# B&R Automation Studio project AS_Project
Automation Studio 6.7.1.5; technology packages: OpcUaCs 6.7.0

## Configuration Config1

CPU 5APC3100.KBU2-000, AutomationRuntime 6.8.1, Build 11.3.0

### Task classes (Cpu.sw)
```
Cyclic#4:
  AltDBExamp <- AltDBExample.prg
Libraries: AltDB, AsTCP, runtime, AsBrStr
```

### Hardware
```
5APC3100_KBU2_000 : 5APC3100.KBU2-000 v2.3.1.0
  Connector IF3:
    AssignedOperatingSystem = ARemb
    ActivateDevice = 1
  Connector IF4:
    AssignedOperatingSystem = ARemb
    ActivateDevice = 1
  Connector IF5:
    AssignedOperatingSystem = ARemb
  Connector IF6:
    AssignedOperatingSystem = ARemb
  Connector IF7:
    AssignedOperatingSystem = ARemb
  Connector IF8:
    AssignedOperatingSystem = ARemb
  ConfigurationID = AltDB_Config1
  Simulation = 1
  ActivateEncryption = 0
  FileDevice1
  FileDeviceName1 = USER
  FileDevicePath1 = USER_PATH
```

### BRRole.brrole - 5APC3100_KBU2_000/AccessAndSecurity/UserRoleSystem/BRRole.brrole
```
Element BR_Anonymous (Type=BRRole)
Element BR_Engineer (Type=BRRole)
Element BR_Observer (Type=BRRole)
Element BR_SafetyAdmin (Type=BRRole)
Element BR_SecurityAdmin (Type=BRRole)
```

- Physical/Config1/5APC3100_KBU2_000/IoMap.iom: same as Physical/Config1/5APC3100_KBU2_000/Cpu.per
- Physical/Config1/5APC3100_KBU2_000/PvMap.vvm: same as Physical/Config1/5APC3100_KBU2_000/Cpu.per
- Safety project (password-protected, skipped)

## Logical view

Binary libraries used (declarations not repeated): operator, runtime, AsIecCon, AsTCP, AsBrStr

### Global.typ - Global data types
```iecst
TYPE
	ReceipeType : 	STRUCT
		price : REAL;				(*recipe price*)
		setTemp : REAL;				(*set temperature*)
		milk : REAL;				(*milk quantity*)
		sugar : REAL;				(*sugar quantity*)
		coffee : REAL;				(*coffee quantity*)
		water : REAL;				(*water quantity*)
	END_STRUCT;
	ParType : 	STRUCT
		receipe : ReceipeType;		(*active recipe parameters*)
	END_STRUCT;
	MainLogicType : 	STRUCT
		par : ParType;				(*parameter structure*)
	END_STRUCT;
END_TYPE
```

### Global.var - Global variables
```iecst
VAR
gMainLogic : MainLogicType;
END_VAR

VAR CONSTANT

END_VAR
```

### Package Logical/Libraries - Global libraries

### Library Logical/Libraries/AltDB (ANSIC, version 1.0.2)
Depends on: AsTCP

#### Types.typ - Exported data types
```iecst
TYPE
	(*Extension type (not part of AsDb): internal diagnostic snapshot of
	a connection, returned by the extension FB dbGetConnState. Exposes
	the state machine of Section 9.2 plus buffering/parsing counters so
	a stuck connection (e.g. permanently ERR_FUB_BUSY) can be diagnosed
	without reading this library's C sources.*)
	AltDBConnStateType : STRUCT
		state				: UINT;		(*CONNSTATE_*, see Priv.var - OPENING/CONNECTING/PRELOGIN/LOGIN/IDLE/EXECUTING/IN_RESULT/BROKEN/FAILED*)
		netStep				: UINT;		(*sub-state of the current network operation (0=send,1=recv)*)
		jobKind				: UINT;		(*JOB_* - which FB currently owns this connection's job, JOB_NONE if idle*)
		locked				: BOOL;		(*TRUE while a job is in progress on this connection*)
		tcpIdent			: UDINT;	(*AsTCP socket identifier, 0 = not opened yet*)
		encoding			: UINT;		(*DBENC_ISO_8859_1 (0) / DBENC_UTF_8 (1)*)
		packetSize			: UINT;		(*negotiated TDS packet size*)
		sendLen				: UDINT;	(*total bytes of the outgoing message currently being sent*)
		sendPos				: UDINT;	(*bytes already handed to TcpSend*)
		tokLen				: UDINT;	(*bytes currently buffered in the de-framed token stream*)
		tokPos				: UDINT;	(*parser read cursor into the token stream*)
		statementActive		: BOOL;		(*TRUE once dbExecuteSql has completed at least once*)
		columnCount			: INT;		(*column count of the current result set, 0 if none*)
		hasResultSet		: BOOL;		(*current statement produced a result set*)
		resultSetOpen		: BOOL;		(*result set still has rows pending / not yet exhausted*)
		rowReady			: BOOL;		(*a row is currently buffered and ready for dbGetData*)
		noMoreRows			: BOOL;		(*end of the current result set has been reached*)
		affectedRows		: UDINT;
		affectedRowsKnown	: BOOL;
		diagCount			: UINT;		(*number of diagnostic records currently in the ring*)
		diagReadIdx			: UINT;		(*index of the next unread diagnostic record*)
		serverVersion		: STRING[31];	(*"mm.mm.bbbb" once LOGINACK has been received, else empty*)
	END_STRUCT;
END_TYPE
```

#### Constants.var - Exported constants
```iecst
VAR CONSTANT
	DB_SYSTEM_SYBASE				: UINT := 1;		(*Sybase database*)
	DB_SYSTEM_MS_SQL				: UINT := 2;		(*Microsoft SQL database*)

	DB_DEFAULT_PORT					: UINT := 5000;		(*default database port*)

	DB_SQL_ERROR					: INT := -1;		(*SQL error*)
	DB_SQL_INVALID_HANDLE			: INT := -2;		(*invalid SQL database handle*)
	DB_SQL_NO_DATA					: INT := 100;		(*no data available*)

	DB_SQL_CHAR						: INT := 1;			(*character data type of either fixed length or variable length*)
	DB_SQL_NUMERIC					: INT := 2;			(*numeric data type with fixed precision and scale*)
	DB_SQL_DECIMAL					: INT := 3;			(*numeric data type with fixed precision and scale*)
	DB_SQL_BIGINT					: INT := -25;		(*big integer 8 bytes*)
	DB_SQL_INTEGER					: INT := 4;			(*DINT*)
	DB_SQL_SMALLINT					: INT := 5;			(*INT*)
	DB_SQL_TINYINT					: INT := -6;		(*SINT*)
	DB_SQL_REAL						: INT := 7;			(*REAL*)
	DB_SQL_DOUBLE					: INT := 8;			(*LREAL*)
	DB_SQL_DATE						: INT := 9;			(*date, 6 bytes: yy.mm.dd*)
	DB_SQL_TIME						: INT := 10;		(*time of a day without time zone based on a 24-hour clock, 6 bytes: hh:mm:ss*)
	DB_SQL_TIMESTAMP				: INT := 11;		(*DB_SQL_DATE + TIME 12 bytes: yy.mm.dd hh:mm:ss*)
	DB_SQL_GUID						: INT := -11;		(*16 byte GUID*)

	DB_IT_SQL_ACCESSIBLE_TABLES				: UINT := 19;		(*SQL_ACCESSIBLE_TABLES*)
	DB_IT_SQL_ACTIVE_ENVIRONMENTS			: UINT := 116;		(*SQL_ACTIVE_ENVIRONMENTS*)
	DB_IT_SQL_AGGREGATE_FUNCTIONS			: UINT := 169;		(*SQL_AGGREGATE_FUNCTIONS*)
	DB_IT_SQL_ALTER_DOMAIN					: UINT := 117;		(*SQL_ALTER_DOMAIN*)
	DB_IT_SQL_ALTER_TABLE					: UINT := 86;		(*SQL_ALTER_TABLE*)
	DB_IT_SQL_ASYNC_MODE					: UINT := 10021;		(*SQL_ASYNC_MODE*)
	DB_IT_SQL_BATCH_ROW_COUNT				: UINT := 120;		(*SQL_BATCH_ROW_COUNT*)
	DB_IT_SQL_BATCH_SUPPORT					: UINT := 121;		(*SQL_BATCH_SUPPORT*)
	DB_IT_SQL_BOOKMARK_PERSISTENCE			: UINT := 82;		(*SQL_BOOKMARK_PERSISTENCE*)
	DB_IT_SQL_CATALOG_LOCATION				: UINT := 114;		(*SQL_CATALOG_LOCATION*)
	DB_IT_SQL_CATALOG_NAME					: UINT := 10003;		(*SQL_CATALOG_NAME*)
	DB_IT_SQL_CATALOG_NAME_SEPARATOR		: UINT := 41;		(*SQL_CATALOG_NAME_SEPARATOR*)
	DB_IT_SQL_CATALOG_TERM					: UINT := 42;		(*SQL_CATALOG_TERM*)
	DB_IT_SQL_CATALOG_USAGE					: UINT := 92;		(*SQL_CATALOG_USAGE*)
	DB_IT_SQL_COLUMN_ALIAS					: UINT := 87;		(*SQL_COLUMN_ALIAS*)
	DB_IT_SQL_CONCAT_NULL_BEHAVIOR			: UINT := 22;		(*SQL_CONCAT_NULL_BEHAVIOR*)
	DB_IT_SQL_CONVERT_BINARY				: UINT := 54;		(*SQL_CONVERT_BINARY*)
	DB_IT_SQL_CONVERT_BIT					: UINT := 55;		(*SQL_CONVERT_BIT*)
	DB_IT_SQL_CONVERT_CHAR					: UINT := 56;		(*SQL_CONVERT_CHAR*)
	DB_IT_SQL_CONVERT_DECIMAL				: UINT := 58;		(*SQL_CONVERT_DECIMAL*)
	DB_IT_SQL_CONVERT_FLOAT					: UINT := 60;		(*SQL_CONVERT_FLOAT*)
	DB_IT_SQL_CONVERT_FUNCTIONS				: UINT := 48;		(*SQL_CONVERT_FUNCTIONS*)
	DB_IT_SQL_CONVERT_INTEGER				: UINT := 61;		(*SQL_CONVERT_INTEGER*)
	DB_IT_SQL_CONVERT_LONGVARBINARY			: UINT := 71;		(*SQL_CONVERT_LONGVARBINARY*)
	DB_IT_SQL_CONVERT_LONGVARCHAR			: UINT := 62;		(*SQL_CONVERT_LONGVARCHAR*)
	DB_IT_SQL_CONVERT_NUMERIC				: UINT := 63;		(*SQL_CONVERT_NUMERIC*)
	DB_IT_SQL_CONVERT_REAL					: UINT := 64;		(*SQL_CONVERT_REAL*)
	DB_IT_SQL_CONVERT_SMALLINT				: UINT := 65;		(*SQL_CONVERT_SMALLINT*)
	DB_IT_SQL_CONVERT_TIMESTAMP				: UINT := 67;		(*SQL_CONVERT_TIMESTAMP*)
	DB_IT_SQL_CONVERT_TINYINT				: UINT := 68;		(*SQL_CONVERT_TINYINT*)
	DB_IT_SQL_CONVERT_VARBINARY				: UINT := 69;		(*SQL_CONVERT_VARBINARY*)
	DB_IT_SQL_CONVERT_VARCHAR				: UINT := 70;		(*SQL_CONVERT_VARCHAR*)
	DB_IT_SQL_CONVERT_WCHAR					: UINT := 122;		(*SQL_CONVERT_WCHAR*)
	DB_IT_SQL_CONVERT_WLONGVARCHAR			: UINT := 125;		(*SQL_CONVERT_WLONGVARCHAR*)
	DB_IT_SQL_CONVERT_WVARCHAR				: UINT := 126;		(*SQL_CONVERT_WVARCHAR*)
	DB_IT_SQL_CORRELATION_NAME				: UINT := 74;		(*SQL_CORRELATION_NAME*)
	DB_IT_SQL_CREATE_ASSERTION				: UINT := 127;		(*SQL_CREATE_ASSERTION*)
	DB_IT_SQL_CREATE_CHARACTER_SET			: UINT := 128;		(*SQL_CREATE_CHARACTER_SET*)
	DB_IT_SQL_CREATE_COLLATION				: UINT := 129;		(*SQL_CREATE_COLLATION*)
	DB_IT_SQL_CREATE_DOMAIN					: UINT := 130;		(*SQL_CREATE_DOMAIN*)
	DB_IT_SQL_CREATE_SCHEMA					: UINT := 131;		(*SQL_CREATE_SCHEMA*)
	DB_IT_SQL_CREATE_TABLE					: UINT := 132;		(*SQL_CREATE_TABLE*)
	DB_IT_SQL_CREATE_TRANSLATION			: UINT := 133;		(*SQL_CREATE_TRANSLATION*)
	DB_IT_SQL_CREATE_VIEW					: UINT := 134;		(*SQL_CREATE_VIEW*)
	DB_IT_SQL_CURSOR_COMMIT_BEHAVIOR		: UINT := 23;		(*SQL_CURSOR_COMMIT_BEHAVIOR*)
	DB_IT_SQL_CURSOR_ROLLBACK_BEHAV			: UINT := 24;		(*SQL_CURSOR_ROLLBACK_BEHAVIOR*)
	DB_IT_SQL_CURSOR_SENSITIVITY			: UINT := 10001;		(*SQL_CURSOR_SENSITIVITY*)
	DB_IT_SQL_DATA_SOURCE_NAME				: UINT := 2;		(*SQL_DATA_SOURCE_NAME*)
	DB_IT_SQL_DATA_SOURCE_READ_ONLY			: UINT := 25;		(*SQL_DATA_SOURCE_READ_ONLY*)
	DB_IT_SQL_DATABASE_NAME					: UINT := 16;		(*SQL_DATABASE_NAME*)
	DB_IT_SQL_DATETIME_LITERALS				: UINT := 119;		(*SQL_DATETIME_LITERALS*)
	DB_IT_SQL_DBMS_NAME						: UINT := 17;		(*SQL_DBMS_NAME*)
	DB_IT_SQL_DBMS_VER						: UINT := 18;		(*SQL_DBMS_VER*)
	DB_IT_SQL_DDL_INDEX						: UINT := 170;		(*SQL_DDL_INDEX*)
	DB_IT_SQL_DEFAULT_TXN_ISOLATION			: UINT := 26;		(*SQL_DEFAULT_TXN_ISOLATION*)
	DB_IT_SQL_DESCRIBE_PARAMETER			: UINT := 10002;		(*SQL_DESCRIBE_PARAMETER*)
	DB_IT_SQL_DRIVER_HDBC					: UINT := 3;		(*SQL_DRIVER_HDBC*)
	DB_IT_SQL_DRIVER_HENV					: UINT := 4;		(*SQL_DRIVER_HENV*)
	DB_IT_SQL_DRIVER_HSTMT					: UINT := 5;		(*SQL_DRIVER_HSTMT*)
	DB_IT_SQL_DRIVER_NAME					: UINT := 6;		(*SQL_DRIVER_NAME*)
	DB_IT_SQL_DRIVER_ODBC_VER				: UINT := 77;		(*SQL_DRIVER_ODBC_VER*)
	DB_IT_SQL_DRIVER_VER					: UINT := 7;		(*SQL_DRIVER_VER*)
	DB_IT_SQL_DROP_ASSERTION				: UINT := 136;		(*SQL_DROP_ASSERTION*)
	DB_IT_SQL_DROP_CHARACTER_SET			: UINT := 137;		(*SQL_DROP_CHARACTER_SET*)
	DB_IT_SQL_DROP_COLLATION				: UINT := 138;		(*SQL_DROP_COLLATION*)
	DB_IT_SQL_DROP_DOMAIN					: UINT := 139;		(*SQL_DROP_DOMAIN*)
	DB_IT_SQL_DROP_SCHEMA					: UINT := 140;		(*SQL_DROP_SCHEMA*)
	DB_IT_SQL_DROP_TABLE					: UINT := 141;		(*SQL_DROP_TABLE*)
	DB_IT_SQL_DROP_TRANSLATION				: UINT := 142;		(*SQL_DROP_TRANSLATION*)
	DB_IT_SQL_DROP_VIEW						: UINT := 143;		(*SQL_DROP_VIEW*)
	DB_IT_SQL_DYNAMIC_CURSOR_ATTR1			: UINT := 144;		(*SQL_DYNAMIC_CURSOR_ATTRIBUTES1*)
	DB_IT_SQL_DYNAMIC_CURSOR_ATTR2			: UINT := 145;		(*SQL_DYNAMIC_CURSOR_ATTRIBUTES2*)
	DB_IT_SQL_EXPRESSIONS_IN_ORDERBY		: UINT := 27;		(*SQL_EXPRESSIONS_IN_ORDERBY*)
	DB_IT_SQL_FETCH_DIRECTION				: UINT := 8;		(*SQL_FETCH_DIRECTION*)
	DB_IT_SQL_FILE_USAGE					: UINT := 84;		(*SQL_FILE_USAGE*)
	DB_IT_SQL_FORW_ONLY_CURSOR_ATTR1		: UINT := 146;		(*SQL_FORWARD_ONLY_CURSOR_ATTRIBUTES1*)
	DB_IT_SQL_FORW_ONLY_CURSOR_ATTR2		: UINT := 147;		(*SQL_FORWARD_ONLY_CURSOR_ATTRIBUTES2*)
	DB_IT_SQL_GETDATA_EXTENSIONS			: UINT := 81;		(*SQL_GETDATA_EXTENSIONS*)
	DB_IT_SQL_GROUP_BY						: UINT := 88;		(*SQL_GROUP_BY*)
	DB_IT_SQL_IDENTIFIER_CASE				: UINT := 28;		(*SQL_IDENTIFIER_CASE*)
	DB_IT_SQL_IDENTIFIER_QUOTE_CHAR			: UINT := 29;		(*SQL_IDENTIFIER_QUOTE_CHAR*)
	DB_IT_SQL_INDEX_KEYWORDS				: UINT := 148;		(*SQL_INDEX_KEYWORDS*)
	DB_IT_SQL_INFO_SCHEMA_VIEWS				: UINT := 149;		(*SQL_INFO_SCHEMA_VIEWS*)
	DB_IT_SQL_INSERT_STATEMENT				: UINT := 172;		(*SQL_INSERT_STATEMENT*)
	DB_IT_SQL_INTEGRITY						: UINT := 73;		(*SQL_INTEGRITY*)
	DB_IT_SQL_KEYSET_CURSOR_ATTR1			: UINT := 150;		(*SQL_KEYSET_CURSOR_ATTRIBUTES1*)
	DB_IT_SQL_KEYSET_CURSOR_ATTR2			: UINT := 151;		(*SQL_KEYSET_CURSOR_ATTRIBUTES2*)
	DB_IT_SQL_KEYWORDS						: UINT := 89;		(*SQL_KEYWORDS*)
	DB_IT_SQL_LIKE_ESCAPE_CLAUSE			: UINT := 113;		(*SQL_LIKE_ESCAPE_CLAUSE*)
	DB_IT_SQL_LOCK_TYPES					: UINT := 78;		(*SQL_LOCK_TYPES*)
	DB_IT_SQL_MAX_ASYNC_CONCUR_STMT			: UINT := 10022;		(*SQL_MAX_ASYNC_CONCURRENT_STATEMENTS*)
	DB_IT_SQL_MAX_BINARY_LITERAL_LEN		: UINT := 112;		(*SQL_MAX_BINARY_LITERAL_LEN*)
	DB_IT_SQL_MAX_CATALOG_NAME_LEN			: UINT := 34;		(*SQL_MAX_CATALOG_NAME_LEN*)
	DB_IT_SQL_MAX_CHAR_LITERAL_LEN			: UINT := 108;		(*SQL_MAX_CHAR_LITERAL_LEN*)
	DB_IT_SQL_MAX_COLUMN_NAME_LEN			: UINT := 30;		(*SQL_MAX_COLUMN_NAME_LEN*)
	DB_IT_SQL_MAX_COLS_IN_GROUP_BY			: UINT := 97;		(*SQL_MAX_COLUMNS_IN_GROUP_BY*)
	DB_IT_SQL_MAX_COLUMNS_IN_INDEX			: UINT := 98;		(*SQL_MAX_COLUMNS_IN_INDEX*)
	DB_IT_SQL_MAX_COLS_IN_ORDER_BY			: UINT := 99;		(*SQL_MAX_COLUMNS_IN_ORDER_BY*)
	DB_IT_SQL_MAX_COLUMNS_IN_SELECT			: UINT := 100;		(*SQL_MAX_COLUMNS_IN_SELECT*)
	DB_IT_SQL_MAX_COLUMNS_IN_TABLE			: UINT := 101;		(*SQL_MAX_COLUMNS_IN_TABLE*)
	DB_IT_SQL_MAX_CONCUR_ACTIVITIES			: UINT := 1;		(*SQL_MAX_CONCURRENT_ACTIVITIES*)
	DB_IT_SQL_MAX_CURSOR_NAME_LEN			: UINT := 31;		(*SQL_MAX_CURSOR_NAME_LEN*)
	DB_IT_SQL_MAX_DRIVER_CONNECTIONS		: UINT := 0;		(*SQL_MAX_DRIVER_CONNECTIONS*)
	DB_IT_SQL_MAX_IDENTIFIER_LEN			: UINT := 10005;		(*SQL_MAX_IDENTIFIER_LEN*)
	DB_IT_SQL_MAX_INDEX_SIZE				: UINT := 102;		(*SQL_MAX_INDEX_SIZE*)
	DB_IT_SQL_MAX_PROCEDURE_NAME_LEN		: UINT := 33;		(*SQL_MAX_PROCEDURE_NAME_LEN*)
	DB_IT_SQL_MAX_ROW_SIZE					: UINT := 104;		(*SQL_MAX_ROW_SIZE*)
	DB_IT_SQL_MAX_ROW_SIZE_INCL_LONG		: UINT := 103;		(*SQL_MAX_ROW_SIZE_INCLUDES_LONG*)
	DB_IT_SQL_MAX_SCHEMA_NAME_LEN			: UINT := 32;		(*SQL_MAX_SCHEMA_NAME_LEN*)
	DB_IT_SQL_MAX_STATEMENT_LEN				: UINT := 105;		(*SQL_MAX_STATEMENT_LEN*)
	DB_IT_SQL_MAX_TABLE_NAME_LEN			: UINT := 35;		(*SQL_MAX_TABLE_NAME_LEN*)
	DB_IT_SQL_MAX_TABLES_IN_SELECT			: UINT := 106;		(*SQL_MAX_TABLES_IN_SELECT*)
	DB_IT_SQL_MAX_USER_NAME_LEN				: UINT := 107;		(*SQL_MAX_USER_NAME_LEN*)
	DB_IT_SQL_MULT_RESULT_SETS				: UINT := 36;		(*SQL_MULT_RESULT_SETS*)
	DB_IT_SQL_MULTIPLE_ACTIVE_TXN			: UINT := 37;		(*SQL_MULTIPLE_ACTIVE_TXN*)
	DB_IT_SQL_NEED_LONG_DATA_LEN			: UINT := 111;		(*SQL_NEED_LONG_DATA_LEN*)
	DB_IT_SQL_NON_NULLABLE_COLUMNS			: UINT := 75;		(*SQL_NON_NULLABLE_COLUMNS*)
	DB_IT_SQL_NULL_COLLATION				: UINT := 85;		(*SQL_NULL_COLLATION*)
	DB_IT_SQL_NUMERIC_FUNCTIONS				: UINT := 49;		(*SQL_NUMERIC_FUNCTIONS*)
	DB_IT_SQL_ODBC_API_CONFORMANCE			: UINT := 9;		(*SQL_ODBC_API_CONFORMANCE*)
	DB_IT_SQL_ODBC_IFC_CONFORMANCE			: UINT := 152;		(*SQL_ODBC_INTERFACE_CONFORMANCE*)
	DB_IT_SQL_ODBC_SAG_CLI_CONFORM			: UINT := 12;		(*SQL_ODBC_SAG_CLI_CONFORMANCE*)
	DB_IT_SQL_ODBC_SQL_CONFORMANCE			: UINT := 15;		(*SQL_ODBC_SQL_CONFORMANCE*)
	DB_IT_SQL_ODBC_VER						: UINT := 10;		(*SQL_ODBC_VER*)
	DB_IT_SQL_OJ_CAPABILITIES				: UINT := 115;		(*SQL_OJ_CAPABILITIES*)
	DB_IT_SQL_ORDER_BY_COLS_IN_SEL			: UINT := 90;		(*SQL_ORDER_BY_COLUMNS_IN_SELECT*)
	DB_IT_SQL_OUTER_JOINS					: UINT := 38;		(*SQL_OUTER_JOINS*)
	DB_IT_SQL_PARAM_ARRAY_ROW_COUNTS		: UINT := 153;		(*SQL_PARAM_ARRAY_ROW_COUNTS*)
	DB_IT_SQL_PARAM_ARRAY_SELECTS			: UINT := 154;		(*SQL_PARAM_ARRAY_SELECTS*)
	DB_IT_SQL_POS_OPERATIONS				: UINT := 79;		(*SQL_POS_OPERATIONS*)
	DB_IT_SQL_POSITIONED_STATEMENTS			: UINT := 80;		(*SQL_POSITIONED_STATEMENTS*)
	DB_IT_SQL_PROCEDURE_TERM				: UINT := 40;		(*SQL_PROCEDURE_TERM*)
	DB_IT_SQL_PROCEDURES					: UINT := 21;		(*SQL_PROCEDURES*)
	DB_IT_SQL_QUOTED_IDENTIFIER_CASE		: UINT := 93;		(*SQL_QUOTED_IDENTIFIER_CASE*)
	DB_IT_SQL_ROW_UPDATES					: UINT := 11;		(*SQL_ROW_UPDATES*)
	DB_IT_SQL_SCHEMA_TERM					: UINT := 39;		(*SQL_SCHEMA_TERM*)
	DB_IT_SQL_SCHEMA_USAGE					: UINT := 91;		(*SQL_SCHEMA_USAGE*)
	DB_IT_SQL_SCROLL_CONCURRENCY			: UINT := 43;		(*SQL_SCROLL_CONCURRENCY*)
	DB_IT_SQL_SCROLL_OPTIONS				: UINT := 44;		(*SQL_SCROLL_OPTIONS*)
	DB_IT_SQL_SEARCH_PATTERN_ESCAPE			: UINT := 14;		(*SQL_SEARCH_PATTERN_ESCAPE*)
	DB_IT_SQL_SERVER_NAME					: UINT := 13;		(*SQL_SERVER_NAME*)
	DB_IT_SQL_SPECIAL_CHARACTERS			: UINT := 94;		(*SQL_SPECIAL_CHARACTERS*)
	DB_IT_SQL_SQL_CONFORMANCE				: UINT := 118;		(*SQL_SQL_CONFORMANCE*)
	DB_IT_SQL_SQL92_DATETIME_FUNCS			: UINT := 155;		(*SQL_SQL92_DATETIME_FUNCTIONS*)
	DB_IT_SQL_SQL92_FK_DELETE_RULE			: UINT := 156;		(*SQL_SQL92_FOREIGN_KEY_DELETE_RULE*)
	DB_IT_SQL_SQL92_FK_UPDATE_RULE			: UINT := 157;		(*SQL_SQL92_FOREIGN_KEY_UPDATE_RULE*)
	DB_IT_SQL_SQL92_GRANT					: UINT := 158;		(*SQL_SQL92_GRANT*)
	DB_IT_SQL_SQL92_NUM_VALUE_FUNCS			: UINT := 159;		(*SQL_SQL92_NUMERIC_VALUE_FUNCTIONS*)
	DB_IT_SQL_SQL92_PREDICATES				: UINT := 160;		(*SQL_SQL92_PREDICATES*)
	DB_IT_SQL_SQL92_REL_JOIN_OPS			: UINT := 161;		(*SQL_SQL92_RELATIONAL_JOIN_OPERATORS*)
	DB_IT_SQL_SQL92_REVOKE					: UINT := 162;		(*SQL_SQL92_REVOKE*)
	DB_IT_SQL_SQL92_ROW_VALUE_CTOR			: UINT := 163;		(*SQL_SQL92_ROW_VALUE_CONSTRUCTOR*)
	DB_IT_SQL_SQL92_STRING_FUNCTIONS		: UINT := 164;		(*SQL_SQL92_STRING_FUNCTIONS*)
	DB_IT_SQL_SQL92_VALUE_EXPR				: UINT := 165;		(*SQL_SQL92_VALUE_EXPRESSIONS*)
	DB_IT_SQL_STD_CLI_CONFORMANCE			: UINT := 166;		(*SQL_STANDARD_CLI_CONFORMANCE*)
	DB_IT_SQL_STATIC_CURSOR_ATTR1			: UINT := 167;		(*SQL_STATIC_CURSOR_ATTRIBUTES1*)
	DB_IT_SQL_STATIC_CURSOR_ATTR2			: UINT := 168;		(*SQL_STATIC_CURSOR_ATTRIBUTES2*)
	DB_IT_SQL_STATIC_SENSITIVITY			: UINT := 83;		(*SQL_STATIC_SENSITIVITY*)
	DB_IT_SQL_STRING_FUNCTIONS				: UINT := 50;		(*SQL_STRING_FUNCTIONS*)
	DB_IT_SQL_SUBQUERIES					: UINT := 95;		(*SQL_SUBQUERIES*)
	DB_IT_SQL_SYSTEM_FUNCTIONS				: UINT := 51;		(*SQL_SYSTEM_FUNCTIONS*)
	DB_IT_SQL_TABLE_TERM					: UINT := 45;		(*SQL_TABLE_TERM*)
	DB_IT_SQL_TIMEDATE_ADD_INTERVALS		: UINT := 109;		(*SQL_TIMEDATE_ADD_INTERVALS*)
	DB_IT_SQL_TIMEDATE_DIFF_INTERVAL		: UINT := 110;		(*SQL_TIMEDATE_DIFF_INTERVALS*)
	DB_IT_SQL_TIMEDATE_FUNCTIONS			: UINT := 52;		(*SQL_TIMEDATE_FUNCTIONS*)
	DB_IT_SQL_TXN_CAPABLE					: UINT := 46;		(*SQL_TXN_CAPABLE*)
	DB_IT_SQL_TXN_ISOLATION_OPTION			: UINT := 72;		(*SQL_TXN_ISOLATION_OPTION*)
	DB_IT_SQL_UNION							: UINT := 96;		(*SQL_UNION*)
	DB_IT_SQL_USER_NAME						: UINT := 47;		(*SQL_USER_NAME*)
	DB_IT_SQL_XOPEN_CLI_YEAR				: UINT := 10000;	(*SQL_XOPEN_CLI_YEAR*)

	dbERR_MEMORY 					: UINT := 34930;	(*memory error*)
	dbERR_DATABASE					: UINT := 34931;	(*database returned an error*)
	dbERR_INVALID_HANDLE			: UINT := 34932;	(*invalid handle specified*)
	dbERR_INVALID_COLUMN			: UINT := 34933;	(*invalid column index specified*)
	dbERR_UNSUPPORTED_DATABASE		: UINT := 34934;	(*unsupported database*)
	dbERR_BUFFER_SIZE				: UINT := 34935;	(*buffer too small*)
	dbERR_INVALID_SERVERNAME		: UINT := 34936;	(*invalid server name*)
	dbERR_INVALID_USERNAME  		: UINT := 34937;	(*invalid user name*)
	dbERR_INVALID_PASSWORD  		: UINT := 34938;	(*invalid password*)
	dbERR_INVALID_DATABASE_NAME 	: UINT := 34939;	(*invalid database name*)
	dbERR_INVALID_SQL_STATEMENT 	: UINT := 34940;	(*invalid SQL statement*)
	dbERR_SQL_EXECUTE_REQUIRED		: UINT := 34941;	(*dbExecuteSql() must be called before*)
	dbERR_INVALID_DATATYPE			: UINT := 34942;	(*invalid data type*)
	dbERR_NULLPOINTER				: UINT := 34943;	(*null pointer*)
	dbERR_NOT_AVAILABLE				: UINT := 34944;	(*information not available*)
	dbERR_UNSUPPORTED_ENCODING		: UINT := 34945;	(*unsupported encoding specified*)
END_VAR

VAR CONSTANT
	DB_ENCODING_ISO_8859_1			: STRING[12] := 'ISO-8859-1';	(*ISO-8859-1 encoding*)
	DB_ENCODING_UTF_8				: STRING[12] := 'UTF-8';		(*UTF-8 encoding*)
END_VAR
```

#### AltDB.fun - Exported functions and function blocks
```iecst
{REDUND_CONTEXT} {REDUND_UNREPLICABLE} FUNCTION_BLOCK dbConnect						(*connects to an existing database; asynchronous execution*)
	VAR_INPUT
		enable			: BOOL;					(*enables execution*)
		pServerName		: UDINT;				(*pointer to IP address or host name of the database server, e.g. "sun.galaxy.one"*)
		pUserName		: UDINT;				(*pointer to the user name*)
		pPassword		: UDINT;				(*pointer to the user password*)
		pDatabaseName	: UDINT;				(*pointer to the name of the database*)
		databaseSystem	: UDINT;				(*database system*)
	END_VAR

	VAR_OUTPUT
		status		 	: UINT;					(*execution status: ERR_OK, ERR_FUB_ENABLE_FALSE, ERR_FUB_BUSY, 0xXXXX = see help*)
		dbError		 	: INT;					(*error number of the database*)
		connectionIdent	: UDINT;				(*identifier of the database connection*)
	END_VAR

	VAR
		_statemachine	: UINT;					(*internal variable*)
		_result			: UINT;					(*internal variable*)
	END_VAR
END_FUNCTION_BLOCK

{REDUND_CONTEXT} {REDUND_UNREPLICABLE} FUNCTION_BLOCK dbConnectEnc						(*connects to an existing database using given encoding; asynchronous execution*)
	VAR_INPUT
		enable			: BOOL;					(*enables execution*)
		pServerName		: UDINT;				(*pointer to IP address or host name of the database server, e.g. "sun.galaxy.one"*)
		pUserName		: UDINT;				(*pointer to the user name*)
		pPassword		: UDINT;				(*pointer to the user password*)
		pDatabaseName	: UDINT;				(*pointer to the name of the database*)
		databaseSystem	: UDINT;				(*database system*)
		pEncoding		: UDINT;				(*character encoding*)
	END_VAR

	VAR_OUTPUT
		status		 	: UINT;					(*execution status: ERR_OK, ERR_FUB_ENABLE_FALSE, ERR_FUB_BUSY, 0xXXXX = see help*)
		dbError		 	: INT;					(*error number of the database*)
		connectionIdent	: UDINT;				(*identifier of the database connection*)
	END_VAR

	VAR
		_statemachine	: UINT;					(*internal variable*)
		_result			: UINT;					(*internal variable*)
	END_VAR
END_FUNCTION_BLOCK

{REDUND_CONTEXT} {REDUND_UNREPLICABLE} FUNCTION_BLOCK dbExecuteSql						(*executes an SQL statement; asynchronous execution*)
	VAR_INPUT
		enable			: BOOL;					(*enables execution*)
		connectionIdent	: UDINT;				(*identifier of the database connection*)
		pSqlStatement	: UDINT;				(*pointer to the SQL statement*)
	END_VAR

	VAR_OUTPUT
		status			: UINT;					(*execution status: ERR_OK, ERR_FUB_ENABLE_FALSE, ERR_FUB_BUSY, 0xXXXX = see help*)
		dbError			: INT;					(*error number of the database*)
	END_VAR

	VAR
		_statemachine	: UINT;					(*internal variable*)
		_result			: UINT;					(*internal variable*)
	END_VAR
END_FUNCTION_BLOCK

{REDUND_CONTEXT} {REDUND_UNREPLICABLE} FUNCTION_BLOCK dbGetAffectedRows				(*determines the number of rows affected by an INSERT, UPDATE or DELETE SQL statement; asynchronous execution*)
	VAR_INPUT
		enable			: BOOL;					(*enables execution*)
		connectionIdent	: UDINT;				(*identifier of the database connection*)
	END_VAR

	VAR_OUTPUT
		status			: UINT;					(*execution status: ERR_OK, ERR_FUB_ENABLE_FALSE, ERR_FUB_BUSY, 0xXXXX = see help*)
		dbError			: INT;					(*error number of the database*)
		affectedRows: UDINT;					(*number of affected rows*)
	END_VAR

	VAR
		_statemachine	: UINT;					(*internal variable*)
		_result			: UINT;					(*internal variable*)
	END_VAR
END_FUNCTION_BLOCK

{REDUND_CONTEXT} {REDUND_UNREPLICABLE} FUNCTION_BLOCK dbGetColumnCount					(*determines the number of columns in the result set of an SELECT SQL statement; asynchronous execution*)
	VAR_INPUT
		enable			: BOOL;					(*enables execution*)
		connectionIdent	: UDINT;				(*identifier of the database connection*)
	END_VAR

	VAR_OUTPUT
		status			: UINT;					(*execution status: ERR_OK, ERR_FUB_ENABLE_FALSE, ERR_FUB_BUSY, 0xXXXX = see help*)
		dbError			: INT;					(*error number of the database*)
		columnCount 	: INT;					(*number of columns in the result set*)
	END_VAR

	VAR
		_statemachine	: UINT;					(*internal variable*)
		_result			: UINT;					(*internal variable*)
	END_VAR
END_FUNCTION_BLOCK

{REDUND_CONTEXT} {REDUND_UNREPLICABLE} FUNCTION_BLOCK dbFetchNextRow					(*fetches the next row into the memory; asynchronous execution*)
	VAR_INPUT
		enable			: BOOL;					(*enables execution*)
		connectionIdent	: UDINT;				(*identifier of the database connection*)
	END_VAR

	VAR_OUTPUT
		status			: UINT;					(*execution status: ERR_OK, ERR_FUB_ENABLE_FALSE, ERR_FUB_BUSY, 0xXXXX = see help*)
		dbError			: INT;					(*error number of the database*)
	END_VAR

	VAR
		_statemachine	: UINT;					(*internal variable*)
		_result			: UINT;					(*internal variable*)
	END_VAR
END_FUNCTION_BLOCK

{REDUND_CONTEXT} {REDUND_UNREPLICABLE} FUNCTION_BLOCK dbGetData						(*gets the data of the current row of the given column*)
	VAR_INPUT
		enable			: BOOL;					(*enables execution*)
		connectionIdent	: UDINT;				(*identifier of the database connection*)
		columnIdx		: UDINT;				(*the data column index*)
		dataType		: INT;					(*type of the data*)
		pData			: UDINT;				(*pointer to the data buffer*)
		dataSize		: UDINT;				(*size of the data buffer*)
	END_VAR

	VAR_OUTPUT
		status			: UINT;					(*execution status: ERR_OK, ERR_FUB_ENABLE_FALSE, ERR_FUB_BUSY, 0xXXXX = see help*)
		dbError			: INT;					(*error number of the database*)
		actDataSize		: UDINT;				(*size of the written data or needed data size*)
	END_VAR
END_FUNCTION_BLOCK

{REDUND_CONTEXT} {REDUND_UNREPLICABLE} FUNCTION_BLOCK dbDisconnect						(*disconnects the connection to the database; asynchronous execution*)
	VAR_INPUT
		enable			: BOOL;					(*enables execution*)
		connectionIdent	: UDINT;				(*identifier of the database connection*)
	END_VAR

	VAR_OUTPUT
		status			: UINT;					(*execution status: ERR_OK, ERR_FUB_ENABLE_FALSE, ERR_FUB_BUSY, 0xXXXX = see help*)
		dbError			: INT;					(*error number of the database*)
	END_VAR

	VAR
		_statemachine	: UINT;					(*internal variable*)
		_result			: UINT;					(*internal variable*)
	END_VAR
END_FUNCTION_BLOCK

{REDUND_CONTEXT} {REDUND_UNREPLICABLE} FUNCTION_BLOCK dbGetInfo						(*gets database information; asynchronous execution*)
	VAR_INPUT
		enable			: BOOL;					(*enables execution*)
		connectionIdent	: UDINT;				(*identifier of the database connection*)
		infoType		: UINT;					(*type of information*)
		pServerInfo		: UDINT;				(*pointer to buffer for the database information*)
		serverInfoSize	: UDINT;				(*size of the buffer*)
	END_VAR

	VAR_OUTPUT
		status			: UINT;					(*execution status: ERR_OK, ERR_FUB_ENABLE_FALSE, ERR_FUB_BUSY, 0xXXXX = see help*)
		dbError			: INT;					(*error number of the database*)
		actServerInfoSize	: UINT;				(*current size of database information or needed size*)
	END_VAR

	VAR
		_statemachine	: UINT;					(*internal variable*)
		_result			: UINT;					(*internal variable*)
	END_VAR
END_FUNCTION_BLOCK

{REDUND_CONTEXT} {REDUND_UNREPLICABLE} FUNCTION_BLOCK dbGetErrorMessage				(*gets the current database error message; asynchronous execution*)
	VAR_INPUT
		enable			: BOOL;					(*enables execution*)
		connectionIdent	: UDINT;				(*identifier of the database connection*)
		pErrorMessage	: UDINT;				(*buffer for the database error message*)
		errorMessageSize: UDINT;				(*size of the buffer*)
	END_VAR

	VAR_OUTPUT
		status			: UINT;					(*execution status: ERR_OK, ERR_FUB_ENABLE_FALSE, ERR_FUB_BUSY, 0xXXXX = see help*)
		dbError			: INT;					(*error number of the database*)
		sqlState		: ARRAY [0..5] OF USINT;(*five-character SQLSTATE code*)
		nativeError		: DINT;					(*native error code, specific to the data source*)
		actErrorMessageSize	: INT;				(*current size for the error message of the database or necessary size*)
	END_VAR

	VAR
		_statemachine	: UINT;					(*internal variable*)
		_result			: UINT;					(*internal variable*)
	END_VAR
END_FUNCTION_BLOCK

{REDUND_CONTEXT} {REDUND_UNREPLICABLE} FUNCTION_BLOCK dbGetConnState				(*extension FB (not part of AsDb): returns an internal diagnostic snapshot of a connection; synchronous execution*)
	VAR_INPUT
		enable			: BOOL;					(*enables execution*)
		connectionIdent	: UDINT;				(*identifier of the database connection*)
	END_VAR

	VAR_OUTPUT
		status			: UINT;					(*execution status: ERR_OK, ERR_FUB_ENABLE_FALSE, ERR_FUB_BUSY, 0xXXXX = see help*)
		dbError			: INT;					(*error number of the database*)
		connState		: AltDBConnStateType;	(*internal diagnostic snapshot, see Types.typ*)
	END_VAR
END_FUNCTION_BLOCK
```

#### Priv.var - Private implementation constants
```iecst
(********************************************************************
 * Library: AltDB
 * File: Priv.var
 ********************************************************************
 * Private (implementation-only) constants.
 * Not part of the AsDb-compatible public interface (see Types.typ,
 * Constants.var and AltDB.fun, which must stay unchanged).
 *
 * Note: a static library in Automation Studio cannot declare its own
 * (non-constant) global VAR - persistent state belongs to the FB
 * instance of the *caller*. The connection pool shared by all FBs of
 * this library (and the AsTCP FB instances it drives) is therefore
 * kept as ordinary C file-scope variables, declared in State.h and
 * defined once in State.c, not as IEC variables. Because this is a
 * Library, _REPLACE_CONST is always active for its own translation
 * units (confirmed by B&R's "Using PLC constants in ANSI C/C++
 * programs" documentation), so the constants below are compiled as
 * real #define's here and may be used in array bounds / switch-case
 * within this library's own *.c files.
 ********************************************************************)

VAR CONSTANT
	MAX_CONN				: UDINT := 8;		(*size of the connection pool, FR-07. Keep in sync with State.h*)
	MAX_COLUMNS				: UDINT := 32;		(*max columns decoded per result set. Keep in sync with State.h*)
	MAX_COL_VALUE_LEN		: UDINT := 512;		(*max raw bytes stored per column value. Keep in sync with State.h*)
	MAX_DIAG				: UDINT := 8;		(*diagnostics ring size per connection. Keep in sync with State.h*)
	TDS_DEFAULT_PACKET_SIZE	: UINT := 4096;
	JOB_ABANDON_TICKS		: UDINT := 150000;	(*watchdog: ~ cycles before an abandoned job is cancelled*)
	SQL_MAX_LEN				: UDINT := 4096;	(*max encoded SQL statement length; a documented reduction from the
												  AsDb default of 65535 because this library sends every request as
												  a single TDS packet (see Net.c / Common.h)*)

	(* connection slot states, Section 9.2 (TLS states omitted, not implemented) *)
	CONNSTATE_FREE			: UINT := 0;
	CONNSTATE_OPENING		: UINT := 1;		(*TcpOpen in progress*)
	CONNSTATE_CONNECTING	: UINT := 2;		(*TcpClient in progress*)
	CONNSTATE_PRELOGIN		: UINT := 3;		(*PRELOGIN sent, awaiting response*)
	CONNSTATE_LOGIN			: UINT := 4;		(*LOGIN7 sent, awaiting LOGINACK/DONE*)
	CONNSTATE_IDLE			: UINT := 5;		(*ready for a batch*)
	CONNSTATE_EXECUTING		: UINT := 6;		(*batch sent, awaiting first result*)
	CONNSTATE_IN_RESULT		: UINT := 7;		(*result set open, rows pending*)
	CONNSTATE_CLOSING		: UINT := 8;		(*TcpClose in progress*)
	CONNSTATE_BROKEN		: UINT := 9;		(*socket/protocol error, only dbDisconnect/dbGetErrorMessage usable*)
	CONNSTATE_FAILED		: UINT := 10;		(*login failed, only dbDisconnect/dbGetErrorMessage usable*)

	(* job kinds - identifies which FB currently owns the connection's async job *)
	JOB_NONE				: UINT := 0;
	JOB_CONNECT				: UINT := 1;
	JOB_EXECUTE				: UINT := 2;
	JOB_FETCH				: UINT := 3;
	JOB_DISCONNECT			: UINT := 4;

	(* connection character encodings *)
	DBENC_ISO_8859_1		: UINT := 0;
	DBENC_UTF_8				: UINT := 1;

	(* connection handle layout, Section 9.1 *)
	HANDLE_TAG				: UDINT := 16#DB000000;
	HANDLE_SLOT_MASK		: UDINT := 16#00000FFF;
	HANDLE_GEN_SHIFT		: UDINT := 12;
END_VAR
```

#### State.h - Internal connection pool data structures (plain C)
```c
/********************************************************************
 * Library: AltDB
 * File: State.h
 ********************************************************************
 * Internal connection pool storage.
 *
 * A static library in Automation Studio cannot declare its own
 * (non-constant) global IEC variable - persistent data belongs to
 * the FB instance of the caller. Since dbExecuteSql/dbFetchNextRow/
 * dbGetData/... must all reach the *same* connection state by
 * connectionIdent regardless of which FB instance (and which task)
 * calls them, and since that state also has to embed AsTCP's own FB
 * instances (TcpOpen/TcpClient/TcpSend/TcpRecv/TcpClose - which, by
 * IEC 61131-3 rules, cannot be nested inside an IEC STRUCT), the
 * connection pool is implemented as a plain hand-written C structure
 * with ordinary (non-static, so it is shared across this library's
 * translation units) file scope storage, defined once in State.c.
 ********************************************************************/
#ifndef _ALTDB_STATE_H_
#define _ALTDB_STATE_H_

#define ND_MAX_CONN            8		/* keep in sync with MAX_CONN in Priv.var */
#define ND_MAX_COLUMNS          32		/* keep in sync with MAX_COLUMNS in Priv.var */
#define ND_MAX_COL_VALUE_LEN   512		/* keep in sync with MAX_COL_VALUE_LEN in Priv.var */
#define ND_MAX_DIAG              8		/* keep in sync with MAX_DIAG in Priv.var */
#define ND_RECV_SCRATCH_SIZE  4096
#define ND_TOK_BUF_SIZE       8192
#define ND_SEND_BUF_SIZE      4352

typedef struct ColumnInfo
{
	unsigned char DataType;		/* raw TDS TYPE_INFO type id */
	UDINT         MaxLength;	/* TYPE_INFO max length, 0xFFFFFFFF = PLP (MAX) type */
	unsigned char Precision;
	unsigned char Scale;
	BOOL          IsUnicode;	/* UTF-16LE source (N-prefixed types) */
	BOOL          IsPlp;		/* partially length prefixed value encoding */
	BOOL          IsLongLen;	/* legacy TEXT/NTEXT/IMAGE value encoding */
	BOOL          Supported;	/* FALSE for types this library cannot decode */
} ColumnInfo;

typedef struct DiagRec
{
	BOOL          Used;
	BOOL          IsError;		/* class >= 11 */
	char          SqlState[6];	/* 5 ASCII chars + NUL */
	DINT          NativeError;
	UINT          MessageLen;
	char          Message[256];	/* NUL-terminated, connection encoding */
} DiagRec;

typedef struct ConnSlot
{
	/* --- lifecycle / handle validation --- */
	UINT   State;			/* CONNSTATE_*, Priv.var */
	UINT   Generation;		/* incremented on free, part of connectionIdent */
	BOOL   Locked;			/* try-lock for FB calls on this connection */
	UINT   JobKind;			/* JOB_*, which operation currently owns the job */
	UDINT  JobOwner;		/* identity of the owning FB instance (its ADR), 0 = none */
	UDINT  JobTicks;		/* watchdog: cycles since job last served */
	BOOL   Abandoned;		/* TRUE if a dbConnect/dbConnectEnc job on this handle was
							   cancelled mid-flight (enable := FALSE while BUSY, Section
							   9.3). The next dbConnect/dbConnectEnc call on this handle
							   re-captures the (possibly corrected) inputs and restarts
							   the handshake from CONNSTATE_OPENING instead of blindly
							   resuming stale state

	/* --- TCP / TDS framing --- */
	UDINT  TcpIdent;		/* 0 = socket not opened */
	UINT   NetStep;			/* sub-state of the current network operation */
	UINT   Encoding;		/* DBENC_ISO_8859_1 / DBENC_UTF_8 */
	UINT   PacketSize;		/* negotiated TDS packet size */

	TcpOpen_typ   tcpOpen;
	TcpClient_typ tcpClient;
	TcpSend_typ   tcpSend;
	TcpRecv_typ   tcpRecv;
	TcpClose_typ  tcpClose;

	/* --- login parameters, copied from the FB inputs at job start --- */
	char   HostBuf[128];		/* NUL-terminated host name / IP, no port */
	UINT   Port;
	char   LoginUser[129];
	UDINT  LoginUserLen;
	char   LoginPass[129];
	UDINT  LoginPassLen;
	char   LoginDb[129];
	UDINT  LoginDbLen;

	unsigned char RecvScratch[ND_RECV_SCRATCH_SIZE];
	unsigned char HeaderBuf[8];
	unsigned char HeaderGot;
	UDINT  FrameRemaining;

	unsigned char TokBuf[ND_TOK_BUF_SIZE];
	UDINT  TokLen;
	UDINT  TokPos;

	unsigned char SendBuf[ND_SEND_BUF_SIZE];
	UDINT  SendLen;
	UDINT  SendPos;

	unsigned char TransactionDescr[8];
	char   ServerVersion[32];	/* NUL-terminated "mm.mm.bbbb" */

	/* --- current statement / result set --- */
	BOOL        StatementActive;	/* dbExecuteSql has completed at least once */
	INT         ColumnCount;
	BOOL        RowOverflow;	/* TRUE if a row exceeded ND_MAX_COL_VALUE_LEN for some column (dbERR_MEMORY) */
	ColumnInfo  Columns[ND_MAX_COLUMNS];
	BOOL        HasResultSet;
	BOOL        ResultSetOpen;
	UDINT       AffectedRows;
	BOOL        AffectedRowsKnown;

	BOOL   RowReady;
	BOOL   NoMoreRows;
	BOOL   ColIsNull[ND_MAX_COLUMNS];
	UDINT  ColValueLen[ND_MAX_COLUMNS];
	unsigned char ColValue[ND_MAX_COLUMNS][ND_MAX_COL_VALUE_LEN];
	BOOL   ColAlreadyRead[ND_MAX_COLUMNS];

	/* --- diagnostics ring (per connection) --- */
	UINT     DiagCount;
	UINT     DiagReadIdx;
	DiagRec  Diag[ND_MAX_DIAG];
} ConnSlot;

extern ConnSlot gConn[ND_MAX_CONN];

#endif /* _ALTDB_STATE_H_ */
```

#### State.c - Internal connection pool storage
```c
/********************************************************************
 * Library: AltDB
 * File: State.c
 ********************************************************************
 * Storage definition for the connection pool (see State.h).
 ********************************************************************/
#include <bur/plctypes.h>
#include <runtime.h>
#include <AsTCP.h>
#include <AltDB.h>
#include "State.h"

ConnSlot gConn[ND_MAX_CONN];
```

#### Common.h - Shared implementation declarations
```c
/********************************************************************
 * Library: AltDB
 * File: Common.h
 ********************************************************************
 * Shared declarations for the implementation (*.c) files of this
 * library. Not part of the public interface.
 *
 * Implementation scope / known deviations from Spec.md (documented
 * here once, referenced from the relevant modules):
 *  - No TLS/TDS 8.0 support. PRELOGIN always advertises
 *    ENCRYPTION = NOT_SUPPORTED. Servers that require encryption
 *    (ENCRYPT=ON/REQUIRED) will be rejected with dbERR_DATABASE.
 *  - Host name resolution is delegated to AsTCP's TcpClient, which
 *    accepts both dotted-decimal addresses and host names.
 *  - ATTENTION (query cancellation) is not implemented. A result set
 *    that is not fully read before the next dbExecuteSql is drained
 *    by continuing to read and discard tokens (not by cancelling the
 *    batch on the wire). enable = FALSE on a busy FB abandons local
 *    job ownership but does not cancel the in-flight server request.
 *  - TDS/row buffers are bounded (see Priv.var): results with more
 *    than MAX_COLUMNS columns or column values larger than
 *    MAX_COL_VALUE_LEN are rejected with dbERR_MEMORY/garbled data
 *    is never produced, but the row is not usable.
 *  - TEXT/NTEXT/IMAGE/SQL_VARIANT/UDT and DATETIMEOFFSET columns are
 *    parsed structurally (to keep the token stream in sync) but are
 *    only partially convertible; see Convert.c.
 ********************************************************************/

#ifndef _ALTDB_COMMON_H_
#define _ALTDB_COMMON_H_

#ifndef TRUE
#define TRUE 1
#endif
#ifndef FALSE
#define FALSE 0
#endif

#include "State.h"

/* ---- token parser result / modes (Token.c) ---- */
#define TOK_NEED_MORE          0
#define TOK_GOT_COLMETADATA    1
#define TOK_GOT_DONE_FINAL     2	/* batch finished, no (more) result sets */
#define TOK_GOT_ROW            3
#define TOK_GOT_EOF            4	/* current result set ended, no more rows */
#define TOK_ERROR              5	/* server error class>=11 or protocol error */
#define TOK_ERROR_MEMORY       6	/* row/column too large for internal buffers (dbERR_MEMORY) */

#define TOKMODE_LOGIN   0	/* awaiting LOGINACK + terminal DONE */
#define TOKMODE_EXEC    1	/* awaiting first COLMETADATA or terminal DONE */
#define TOKMODE_FETCH   2	/* awaiting next ROW or end of this result set */
#define TOKMODE_DRAIN   3	/* discard everything up to terminal DONE */

/* ---- network step results (Net.c) ---- */
#define NET_IN_PROGRESS 0
#define NET_DONE        1
#define NET_ERROR       2

/* Util.c */
UDINT  AltDB_MakeHandle(UDINT slot, UINT generation);
BOOL   AltDB_SlotFromHandle(UDINT handle, UDINT *pSlot, UINT *pGeneration);
void   AltDB_SlotReset(UDINT slot);
BOOL   AltDB_SlotAlloc(UDINT *pSlot);
BOOL   AltDB_TryLock(UDINT slot, UDINT owner);
void   AltDB_Unlock(UDINT slot);
BOOL   AltDB_IsOwner(UDINT slot, UDINT owner);

void   AltDB_DiagClear(UDINT slot);
void   AltDB_DiagPushServer(UDINT slot, BOOL isError, DINT nativeError,
                               const char *sqlState, const unsigned char *text, UDINT textLen);
void   AltDB_DiagPushClient(UDINT slot, const char *sqlState, const char *text);

UINT   AltDB_ReadLE16(const unsigned char *p);
UDINT  AltDB_ReadLE32(const unsigned char *p);
unsigned long long AltDB_ReadLE64(const unsigned char *p);
UDINT  AltDB_ReadBE16(const unsigned char *p);
void   AltDB_WriteLE16(unsigned char *p, UINT v);
void   AltDB_WriteLE32(unsigned char *p, UDINT v);
void   AltDB_WriteBE16(unsigned char *p, UINT v);

UDINT  AltDB_EncodeToWire(UINT encoding, const char *src, UDINT srcLen, unsigned char *dst, UDINT dstCap);
UDINT  AltDB_WireToConn(UINT encoding, const unsigned char *src, UDINT srcBytes, unsigned char *dst, UDINT dstCap);
UDINT  AltDB_Utf16leToConn(UINT encoding, const unsigned char *src, UDINT srcBytes, unsigned char *dst, UDINT dstCap);
UDINT  AltDB_ConnToUtf16le(UINT encoding, const unsigned char *src, UDINT srcLen, unsigned char *dst, UDINT dstCap);

UDINT  AltDB_FormatI64(long long v, char *dst, UDINT dstCap);
UDINT  AltDB_FormatDouble(double v, int sigDigits, char *dst, UDINT dstCap);
UDINT  AltDB_FormatDecimal(const unsigned char *magnitude, UDINT magLen, BOOL positive, USINT scale, char *dst, UDINT dstCap);

/* Net.c */
INT    AltDB_NetConnectStep(UDINT slot);
INT    AltDB_NetSendStep(UDINT slot);
INT    AltDB_NetRecvPump(UDINT slot);
INT    AltDB_NetDisconnectStep(UDINT slot);
void   AltDB_BuildPrelogin(UDINT slot);
BOOL   AltDB_BuildLogin7(UDINT slot, const char *user, const char *pass, const char *db, const char *server);
BOOL   AltDB_BuildSqlBatch(UDINT slot, const char *sql, UDINT sqlLen);

/* Token.c */
INT    AltDB_TokenStep(UDINT slot, UINT mode);

/* Convert.c */
void   AltDB_GetData(UDINT slot, UDINT columnIdx, INT dataType, UDINT pData, UDINT dataSize,
                        UINT *status, INT *dbError, UDINT *actDataSize);

#endif /* _ALTDB_COMMON_H_ */
```

#### Util.c - Shared helper routines
```c
/********************************************************************
 * Library: AltDB
 * File: Util.c
 ********************************************************************
 * Shared helpers: connection handle encode/decode, slot pool
 * management, diagnostics ring, byte order helpers, character set
 * transcoding and number formatting for DB_SQL_CHAR output.
 ********************************************************************/
#include <bur/plctypes.h>
#include <runtime.h>
#include <AsTCP.h>
#include <AltDB.h>
#include "Common.h"
#include <string.h>

UDINT AltDB_MakeHandle(UDINT slot, UINT generation)
{
	return HANDLE_TAG | (((UDINT)generation << HANDLE_GEN_SHIFT) & 0xFFFFF000UL) | ((slot + 1) & HANDLE_SLOT_MASK);
}

BOOL AltDB_SlotFromHandle(UDINT handle, UDINT *pSlot, UINT *pGeneration)
{
	UDINT slot;
	UINT generation;

	if ((handle & 0xFF000000UL) != HANDLE_TAG) {
		return FALSE;
	}
	slot = (handle & HANDLE_SLOT_MASK);
	if (slot == 0 || slot > MAX_CONN) {
		return FALSE;
	}
	slot = slot - 1;
	generation = (UINT)((handle >> HANDLE_GEN_SHIFT) & 0x0FFF);
	if (gConn[slot].State == CONNSTATE_FREE || gConn[slot].Generation != generation) {
		return FALSE;
	}
	*pSlot = slot;
	*pGeneration = generation;
	return TRUE;
}

void AltDB_SlotReset(UDINT slot)
{
	UINT keepGeneration = gConn[slot].Generation;

	memset(&gConn[slot], 0, sizeof(gConn[slot]));
	gConn[slot].Generation = keepGeneration;
	gConn[slot].State = CONNSTATE_FREE;
	gConn[slot].PacketSize = TDS_DEFAULT_PACKET_SIZE;
}

BOOL AltDB_SlotAlloc(UDINT *pSlot)
{
	UDINT i;

	for (i = 0; i < MAX_CONN; i++) {
		if (gConn[i].State == CONNSTATE_FREE) {
			AltDB_SlotReset(i);
			*pSlot = i;
			return TRUE;
		}
	}
	return FALSE;
}

BOOL AltDB_TryLock(UDINT slot, UDINT owner)
{
	if (gConn[slot].Locked && gConn[slot].JobOwner != owner) {
		return FALSE;
	}
	gConn[slot].Locked = TRUE;
	gConn[slot].JobOwner = owner;
	return TRUE;
}

void AltDB_Unlock(UDINT slot)
{
	gConn[slot].Locked = FALSE;
	gConn[slot].JobOwner = 0;
	gConn[slot].JobKind = JOB_NONE;
	gConn[slot].JobTicks = 0;
}

BOOL AltDB_IsOwner(UDINT slot, UDINT owner)
{
	return (gConn[slot].Locked && gConn[slot].JobOwner == owner);
}

/* ---------------- diagnostics ring ---------------- */

void AltDB_DiagClear(UDINT slot)
{
	gConn[slot].DiagCount = 0;
	gConn[slot].DiagReadIdx = 0;
	memset(gConn[slot].Diag, 0, sizeof(gConn[slot].Diag));
}

static DiagRec *DiagNextSlot(UDINT slot)
{
	UINT idx;

	if (gConn[slot].DiagCount >= MAX_DIAG) {
		/* ring full: drop the oldest unread record to make room */
		memmove(&gConn[slot].Diag[0], &gConn[slot].Diag[1], sizeof(DiagRec) * (MAX_DIAG - 1));
		idx = (UINT)(MAX_DIAG - 1);
		if (gConn[slot].DiagReadIdx > 0) {
			gConn[slot].DiagReadIdx--;
		}
	} else {
		idx = gConn[slot].DiagCount;
		gConn[slot].DiagCount++;
	}
	return &gConn[slot].Diag[idx];
}

void AltDB_DiagPushServer(UDINT slot, BOOL isError, DINT nativeError,
                             const char *sqlState, const unsigned char *text, UDINT textLen)
{
	DiagRec *rec = DiagNextSlot(slot);
	const char *prefix = "[AltDB][SQL Server]";
	UDINT prefixLen = (UDINT)strlen(prefix);
	UDINT cap = (UDINT)sizeof(rec->Message) - 1;
	UDINT n;

	rec->Used = TRUE;
	rec->IsError = isError;
	rec->NativeError = nativeError;
	memcpy(rec->SqlState, sqlState, 5);
	rec->SqlState[5] = 0;

	n = (prefixLen < cap) ? prefixLen : cap;
	memcpy(rec->Message, prefix, n);
	if (n < cap && textLen > 0) {
		UDINT remain = cap - n;
		UDINT copyLen = (textLen < remain) ? textLen : remain;
		memcpy(&rec->Message[n], text, copyLen);
		n += copyLen;
	}
	rec->Message[n] = 0;
	rec->MessageLen = (UINT)n;
}

void AltDB_DiagPushClient(UDINT slot, const char *sqlState, const char *text)
{
	DiagRec *rec = DiagNextSlot(slot);
	UDINT cap = (UDINT)sizeof(rec->Message) - 1;
	UDINT n;

	rec->Used = TRUE;
	rec->IsError = TRUE;
	rec->NativeError = 0;
	memcpy(rec->SqlState, sqlState, 5);
	rec->SqlState[5] = 0;

	n = (UDINT)strlen(text);
	if (n > cap) {
		n = cap;
	}
	memcpy(rec->Message, "[AltDB]", 9);
	if (9 + n > cap) {
		n = cap - 9;
	}
	memcpy(&rec->Message[9], text, n);
	rec->Message[9 + n] = 0;
	rec->MessageLen = (UINT)(9 + n);
}

/* ---------------- byte order ---------------- */

UINT AltDB_ReadLE16(const unsigned char *p)
{
	return (UINT)(p[0] | (p[1] << 8));
}

UDINT AltDB_ReadLE32(const unsigned char *p)
{
	return (UDINT)p[0] | ((UDINT)p[1] << 8) | ((UDINT)p[2] << 16) | ((UDINT)p[3] << 24);
}

unsigned long long AltDB_ReadLE64(const unsigned char *p)
{
	unsigned long long lo = AltDB_ReadLE32(p);
	unsigned long long hi = AltDB_ReadLE32(p + 4);
	return lo | (hi << 32);
}

UDINT AltDB_ReadBE16(const unsigned char *p)
{
	return (UDINT)((p[0] << 8) | p[1]);
}

void AltDB_WriteLE16(unsigned char *p, UINT v)
{
	p[0] = (unsigned char)(v & 0xFF);
	p[1] = (unsigned char)((v >> 8) & 0xFF);
}

void AltDB_WriteLE32(unsigned char *p, UDINT v)
{
	p[0] = (unsigned char)(v & 0xFF);
	p[1] = (unsigned char)((v >> 8) & 0xFF);
	p[2] = (unsigned char)((v >> 16) & 0xFF);
	p[3] = (unsigned char)((v >> 24) & 0xFF);
}

void AltDB_WriteBE16(unsigned char *p, UINT v)
{
	p[0] = (unsigned char)((v >> 8) & 0xFF);
	p[1] = (unsigned char)(v & 0xFF);
}

/* ---------------- character set transcoding ---------------- */
/* Connection encoding is either ISO-8859-1 (1 byte per code point,
 * identical to Unicode code points U+0000..U+00FF) or UTF-8. Server
 * strings are exchanged as UTF-16LE. Unmappable characters become
 * '?' (Section 11.3/11.4, [V-18]). */

UDINT AltDB_Utf16leToConn(UINT encoding, const unsigned char *src, UDINT srcBytes, unsigned char *dst, UDINT dstCap)
{
	UDINT si = 0;
	UDINT di = 0;

	while (si + 2 <= srcBytes) {
		UINT cp = AltDB_ReadLE16(&src[si]);
		si += 2;

		if (cp >= 0xD800 && cp <= 0xDBFF && si + 2 <= srcBytes) {
			UINT lo = AltDB_ReadLE16(&src[si]);
			if (lo >= 0xDC00 && lo <= 0xDFFF) {
				si += 2;
				cp = 0xFFFD; /* surrogate pair: not representable in 8-bit encodings, replacement char */
			}
		}

		if (encoding == DBENC_UTF_8) {
			if (cp < 0x80) {
				if (di + 1 > dstCap) break;
				dst[di++] = (unsigned char)cp;
			} else if (cp < 0x800) {
				if (di + 2 > dstCap) break;
				dst[di++] = (unsigned char)(0xC0 | (cp >> 6));
				dst[di++] = (unsigned char)(0x80 | (cp & 0x3F));
			} else {
				if (di + 3 > dstCap) break;
				dst[di++] = (unsigned char)(0xE0 | (cp >> 12));
				dst[di++] = (unsigned char)(0x80 | ((cp >> 6) & 0x3F));
				dst[di++] = (unsigned char)(0x80 | (cp & 0x3F));
			}
		} else {
			if (di + 1 > dstCap) break;
			dst[di++] = (cp <= 0xFF) ? (unsigned char)cp : (unsigned char)'?';
		}
	}
	return di;
}

UDINT AltDB_ConnToUtf16le(UINT encoding, const unsigned char *src, UDINT srcLen, unsigned char *dst, UDINT dstCap)
{
	UDINT si = 0;
	UDINT di = 0;

	while (si < srcLen) {
		UINT cp;

		if (encoding == DBENC_UTF_8) {
			unsigned char b0 = src[si];
			if (b0 < 0x80) {
				cp = b0; si += 1;
			} else if ((b0 & 0xE0) == 0xC0 && si + 1 < srcLen) {
				cp = ((b0 & 0x1F) << 6) | (src[si + 1] & 0x3F); si += 2;
			} else if ((b0 & 0xF0) == 0xE0 && si + 2 < srcLen) {
				cp = ((b0 & 0x0F) << 12) | ((src[si + 1] & 0x3F) << 6) | (src[si + 2] & 0x3F); si += 3;
			} else {
				cp = '?'; si += 1;
			}
		} else {
			cp = src[si]; si += 1;
		}

		if (di + 2 > dstCap) break;
		AltDB_WriteLE16(&dst[di], (UINT)cp);
		di += 2;
	}
	return di;
}

UDINT AltDB_EncodeToWire(UINT encoding, const char *src, UDINT srcLen, unsigned char *dst, UDINT dstCap)
{
	return AltDB_ConnToUtf16le(encoding, (const unsigned char *)src, srcLen, dst, dstCap);
}

UDINT AltDB_WireToConn(UINT encoding, const unsigned char *src, UDINT srcBytes, unsigned char *dst, UDINT dstCap)
{
	return AltDB_Utf16leToConn(encoding, src, srcBytes, dst, dstCap);
}

/* ---------------- number formatting (Section 11.3) ---------------- */

UDINT AltDB_FormatI64(long long v, char *dst, UDINT dstCap)
{
	char tmp[24];
	UDINT n = 0;
	BOOL neg = (v < 0);
	unsigned long long u;
	UDINT i;

	u = neg ? (unsigned long long)(-(v + 1)) + 1ULL : (unsigned long long)v;
	do {
		tmp[n++] = (char)('0' + (u % 10ULL));
		u /= 10ULL;
	} while (u != 0 && n < sizeof(tmp));

	i = 0;
	if (neg) {
		if (i >= dstCap) return 0;
		dst[i++] = '-';
	}
	while (n > 0 && i < dstCap) {
		dst[i++] = tmp[--n];
	}
	if (i < dstCap) dst[i] = 0;
	return i;
}

/* Formats an unsigned big integer given as a little-endian byte
 * array (TDS DECIMALN/NUMERICN magnitude) as a decimal string with
 * the given number of fractional digits (scale). */
UDINT AltDB_FormatDecimal(const unsigned char *magnitude, UDINT magLen, BOOL positive, USINT scale, char *dst, UDINT dstCap)
{
	unsigned char num[16];
	char digits[40];
	UDINT nDigits = 0;
	UDINT i;
	UDINT di;
	BOOL allZero;
	BOOL valueIsZero = TRUE;

	if (magLen > sizeof(num)) magLen = sizeof(num);
	memcpy(num, magnitude, magLen);
	for (i = 0; i < magLen; i++) {
		if (num[i] != 0) { valueIsZero = FALSE; break; }
	}

	do {
		UDINT rem = 0;
		allZero = TRUE;
		for (i = magLen; i > 0; i--) {
			UDINT cur = (rem << 8) | num[i - 1];
			num[i - 1] = (unsigned char)(cur / 10);
			if (num[i - 1] != 0) allZero = FALSE;
			rem = cur % 10;
		}
		digits[nDigits++] = (char)('0' + rem);
	} while (!allZero && nDigits < sizeof(digits));

	while (nDigits <= scale && nDigits < sizeof(digits)) {
		digits[nDigits++] = '0';
	}

	di = 0;
	if (!positive && !valueIsZero) {
		if (di < dstCap) dst[di++] = '-';
	}
	for (i = 0; i < nDigits - scale; i++) {
		if (di < dstCap) dst[di++] = digits[nDigits - 1 - i];
	}
	if (scale > 0) {
		if (di < dstCap) dst[di++] = '.';
		for (i = 0; i < scale; i++) {
			if (di < dstCap) dst[di++] = digits[scale - 1 - i];
		}
	}
	if (di < dstCap) dst[di] = 0;
	return di;
}

/* Simple significant-digit formatter for REAL/DOUBLE source values.
 * Not a byte-exact match for the original AsDb/ODBC formatting
 * ([V-14], requires golden capture); produces a correct, readable
 * decimal or exponential representation. */
UDINT AltDB_FormatDouble(double v, int sigDigits, char *dst, UDINT dstCap)
{
	UDINT di = 0;
	BOOL neg = FALSE;
	int exp10 = 0;
	double mant;
	unsigned long long scaled;
	char digits[20];
	int i;
	double scale;

	if (v != v) { /* NaN */
		if (dstCap > 3) { dst[0] = 'N'; dst[1] = 'a'; dst[2] = 'N'; dst[3] = 0; return 3; }
		return 0;
	}
	if (v < 0.0) { neg = TRUE; v = -v; }

	if (v == 0.0) {
		if (dstCap > 1) { dst[0] = '0'; dst[1] = 0; return 1; }
		return 0;
	}

	mant = v;
	while (mant >= 10.0 && exp10 < 60) { mant /= 10.0; exp10++; }
	while (mant < 1.0 && exp10 > -60) { mant *= 10.0; exp10--; }

	scale = 1.0;
	for (i = 1; i < sigDigits; i++) scale *= 10.0;
	scaled = (unsigned long long)(mant * scale + 0.5);

	/* rounding may have produced one extra digit (e.g. 9.999->10.00) */
	{
		unsigned long long maxVal = 1;
		for (i = 0; i < sigDigits; i++) maxVal *= 10ULL;
		if (scaled >= maxVal) { scaled /= 10ULL; exp10++; }
	}

	for (i = sigDigits - 1; i >= 0; i--) {
		digits[i] = (char)('0' + (scaled % 10ULL));
		scaled /= 10ULL;
	}

	if (neg && di < dstCap) dst[di++] = '-';

	if (exp10 < -4 || exp10 >= sigDigits) {
		/* exponential form d.ddddE+nn */
		if (di < dstCap) dst[di++] = digits[0];
		if (sigDigits > 1) {
			if (di < dstCap) dst[di++] = '.';
			for (i = 1; i < sigDigits; i++) {
				if (di < dstCap) dst[di++] = digits[i];
			}
		}
		if (di < dstCap) dst[di++] = 'E';
		if (di < dstCap) dst[di++] = (exp10 >= 0) ? '+' : '-';
		{
			int ae = (exp10 >= 0) ? exp10 : -exp10;
			char ebuf[8];
			int en = 0;
			do { ebuf[en++] = (char)('0' + (ae % 10)); ae /= 10; } while (ae != 0);
			while (en > 0) { if (di < dstCap) dst[di++] = ebuf[--en]; }
		}
	} else if (exp10 >= 0) {
		for (i = 0; i <= exp10; i++) {
			if (di < dstCap) dst[di++] = (i < sigDigits) ? digits[i] : '0';
		}
		if (exp10 + 1 < sigDigits) {
			if (di < dstCap) dst[di++] = '.';
			for (i = exp10 + 1; i < sigDigits; i++) {
				if (di < dstCap) dst[di++] = digits[i];
			}
		}
	} else {
		if (di < dstCap) dst[di++] = '0';
		if (di < dstCap) dst[di++] = '.';
		for (i = 0; i < -exp10 - 1; i++) {
			if (di < dstCap) dst[di++] = '0';
		}
		for (i = 0; i < sigDigits; i++) {
			if (di < dstCap) dst[di++] = digits[i];
		}
	}

	if (di < dstCap) dst[di] = 0;
	return di;
}
```

#### Net.c - TCP/TDS network pump, PRELOGIN and LOGIN7
```c
/********************************************************************
 * Library: AltDB
 * File: Net.c
 ********************************************************************
 * TCP transport (driving AsTCP's TcpOpen/TcpClient/TcpSend/TcpRecv/
 * TcpClose asynchronous function blocks from C), TDS packet framing,
 * PRELOGIN and LOGIN7 message construction.
 *
 * Every outgoing message (PRELOGIN, LOGIN7, SQL batch) is built as a
 * single TDS packet (8-byte header + payload) in SendBuf; see
 * Common.h for the resulting, documented limit on SQL statement
 * length (SQL_MAX_LEN).
 ********************************************************************/
#include <bur/plctypes.h>
#include <runtime.h>
#include <AsTCP.h>
#include <AltDB.h>
#include "Common.h"
#include <string.h>

#define NETSTEP_SEND 0
#define NETSTEP_RECV 1

/* ---------------- TCP driving ---------------- */

static INT PumpTcpOpen(UDINT slot)
{
	TcpOpen_typ *p = &gConn[slot].tcpOpen;

	p->enable = TRUE;
	p->pIfAddr = 0;
	p->port = 0;
	p->options = 0;
	TcpOpen(p);
	if (p->status == ERR_FUB_BUSY) return NET_IN_PROGRESS;
	if (p->status == ERR_OK) {
		gConn[slot].TcpIdent = p->ident;
		return NET_DONE;
	}
	AltDB_DiagPushClient(slot, "08001", "unable to open local TCP socket");
	return NET_ERROR;
}

static INT PumpTcpClient(UDINT slot)
{
	TcpClient_typ *p = &gConn[slot].tcpClient;

	p->enable = TRUE;
	p->ident = gConn[slot].TcpIdent;
	p->pServer = (UDINT)(UDINT)&gConn[slot].HostBuf[0];
	p->portserv = gConn[slot].Port;
	TcpClient(p);
	if (p->status == ERR_FUB_BUSY) return NET_IN_PROGRESS;
	if (p->status == ERR_OK) return NET_DONE;
	AltDB_DiagPushClient(slot, "08001", "TCP connect to server failed");
	return NET_ERROR;
}

INT AltDB_NetSendStep(UDINT slot)
{
	TcpSend_typ *p = &gConn[slot].tcpSend;
	ConnSlot *c = &gConn[slot];

	if (c->SendPos >= c->SendLen) return NET_DONE;

	p->enable = TRUE;
	p->ident = c->TcpIdent;
	p->pData = (UDINT)&c->SendBuf[c->SendPos];
	p->datalen = c->SendLen - c->SendPos;
	p->flags = 0;
	TcpSend(p);
	if (p->status == ERR_FUB_BUSY) return NET_IN_PROGRESS;
	if (p->status == ERR_OK) {
		c->SendPos += p->sentlen;
		return (c->SendPos >= c->SendLen) ? NET_DONE : NET_IN_PROGRESS;
	}
	AltDB_DiagPushClient(slot, "08S01", "TCP send failed, connection lost");
	return NET_ERROR;
}

/* Reads any bytes currently available, strips TDS packet headers and
 * appends the logical payload bytes to TokBuf. Returns the number of
 * new logical bytes appended (0 = nothing available right now, a
 * normal/expected result, not an error), or -1 on a hard socket
 * error. */
INT AltDB_NetRecvPump(UDINT slot)
{
	ConnSlot *c = &gConn[slot];
	TcpRecv_typ *p = &gConn[slot].tcpRecv;
	UDINT produced = 0;
	UDINT si;
	UDINT avail;

	/* compact TokBuf if the parser has already consumed a large prefix */
	if (c->TokPos > 0 && (c->TokPos == c->TokLen || c->TokPos > (UDINT)sizeof(c->TokBuf) / 2)) {
		if (c->TokPos < c->TokLen) {
			memmove(&c->TokBuf[0], &c->TokBuf[c->TokPos], c->TokLen - c->TokPos);
		}
		c->TokLen -= c->TokPos;
		c->TokPos = 0;
	}

	if (c->TokLen >= sizeof(c->TokBuf)) {
		/* parser is not keeping up with a bound buffer; stall receiving */
		return 0;
	}

	p->enable = TRUE;
	p->ident = c->TcpIdent;
	p->pData = (UDINT)&c->RecvScratch[0];
	p->datamax = sizeof(c->RecvScratch);
	p->flags = 0;
	TcpRecv(p);

	if (p->status == ERR_FUB_BUSY) return 0;
	if (p->status != ERR_OK) {
		if (p->status == tcpERR_NO_DATA || p->status == tcpERR_WOULDBLOCK) return 0;
		AltDB_DiagPushClient(slot, "08S01", "TCP receive failed, connection lost");
		return -1;
	}
	avail = p->recvlen;
	if (avail == 0) return 0;

	si = 0;
	while (si < avail) {
		if (c->HeaderGot < 8) {
			UDINT need = 8 - c->HeaderGot;
			UDINT take = (avail - si < need) ? (avail - si) : need;
			memcpy(&c->HeaderBuf[c->HeaderGot], &c->RecvScratch[si], take);
			c->HeaderGot += (USINT)take;
			si += take;
			if (c->HeaderGot < 8) break; /* header itself split across reads */
			c->FrameRemaining = AltDB_ReadBE16(&c->HeaderBuf[2]) - 8;
		}
		{
			UDINT take = avail - si;
			if (take > c->FrameRemaining) take = c->FrameRemaining;
			if (c->TokLen + take > sizeof(c->TokBuf)) {
				take = sizeof(c->TokBuf) - c->TokLen;
			}
			if (take > 0) {
				memcpy(&c->TokBuf[c->TokLen], &c->RecvScratch[si], take);
				c->TokLen += take;
				produced += take;
				si += take;
				c->FrameRemaining -= take;
			}
			if (c->FrameRemaining == 0) {
				c->HeaderGot = 0; /* ready for next physical packet header */
			} else {
				/* buffer pressure: stop for this call, resume next pump */
				break;
			}
		}
	}
	return (INT)produced;
}

INT AltDB_NetDisconnectStep(UDINT slot)
{
	ConnSlot *c = &gConn[slot];
	TcpClose_typ *p = &gConn[slot].tcpClose;

	if (c->TcpIdent == 0) return NET_DONE;

	p->enable = TRUE;
	p->ident = c->TcpIdent;
	p->how = 0;
	TcpClose(p);
	if (p->status == ERR_FUB_BUSY) return NET_IN_PROGRESS;
	c->TcpIdent = 0;
	return NET_DONE;
}

/* ---------------- PRELOGIN ---------------- */

/* PRELOGIN option table: VERSION(6), ENCRYPTION(1), INSTOPT(1),
 * THREADID(4), MARS(1), terminator. Identical layout for request and
 * response (Section 10.3). */
void AltDB_BuildPrelogin(UDINT slot)
{
	ConnSlot *c = &gConn[slot];
	unsigned char *b = c->SendBuf;
	UDINT payloadLen = 26 + 6 + 1 + 1 + 4 + 1; /* 39 */
	UDINT total = 8 + payloadLen;

	memset(b, 0, 8 + payloadLen);
	b[0] = 0x12; b[1] = 0x01; /* type PRELOGIN, status EOM */
	AltDB_WriteBE16(&b[2], (UINT)total);
	b[4] = 0; b[5] = 0; b[6] = 1; b[7] = 0;

	{
		unsigned char *p = &b[8];
		UINT off = 26;

		p[0] = 0x00; AltDB_WriteBE16(&p[1], off); AltDB_WriteBE16(&p[3], 6); off += 6;
		p[5] = 0x01; AltDB_WriteBE16(&p[6], off); AltDB_WriteBE16(&p[8], 1); off += 1;
		p[10] = 0x02; AltDB_WriteBE16(&p[11], off); AltDB_WriteBE16(&p[13], 1); off += 1;
		p[15] = 0x03; AltDB_WriteBE16(&p[16], off); AltDB_WriteBE16(&p[18], 4); off += 4;
		p[20] = 0x04; AltDB_WriteBE16(&p[21], off); AltDB_WriteBE16(&p[23], 1); off += 1;
		p[25] = 0xFF;

		p[26] = 0x0F; p[27] = 0x00; p[28] = 0x00; p[29] = 0x00; p[30] = 0x00; p[31] = 0x00; /* VERSION */
		p[32] = 0x02; /* ENCRYPTION = NOT_SUPPORTED (no TLS in this library) */
		p[33] = 0x00; /* INSTOPT = none */
		p[34] = 0x00; p[35] = 0x00; p[36] = 0x00; p[37] = 0x00; /* THREADID */
		p[38] = 0x00; /* MARS = off */
	}

	c->SendLen = total;
	c->SendPos = 0;
}

/* Parses a buffered PRELOGIN response from TokBuf[TokPos..TokLen).
 * Returns 1 if parsed (TokPos advanced past it), 0 if more bytes are
 * needed, -1 on an unsupported/invalid response (diagnostic pushed). */
static INT ParsePreloginResponse(UDINT slot)
{
	ConnSlot *c = &gConn[slot];
	const unsigned char *b = &c->TokBuf[c->TokPos];
	UDINT avail = c->TokLen - c->TokPos;
	UDINT i;
	UDINT tableLen = 0;
	UDINT dataEnd = 0;
	BOOL haveEncryption = FALSE;
	USINT encryptionVal = 0;

	for (i = 0; ; i += 5) {
		if (i + 1 > avail) return 0;
		if (b[i] == 0xFF) { tableLen = i + 1; break; }
		if (i + 5 > avail) return 0;
		{
			UINT tokOff = (UINT)AltDB_ReadBE16(&b[i + 1]);
			UINT tokLen = (UINT)AltDB_ReadBE16(&b[i + 3]);
			UDINT end = (UDINT)tokOff + (UDINT)tokLen;

			if (end > dataEnd) dataEnd = end;
			if (b[i] == 0x01 && tokLen >= 1) {
				if ((UDINT)tokOff + 1 > avail) return 0; /* ENCRYPTION byte not buffered yet */
				haveEncryption = TRUE;
				encryptionVal = b[tokOff];
			}
		}
		if (i > 200) { AltDB_DiagPushClient(slot, "08001", "malformed PRELOGIN response"); return -1; }
	}

	/* Wait for every byte referenced by the option table (not a fixed
	 * padding guess - SQL Server's PRELOGIN response is tightly sized
	 * with no slack, so an inexact bound here would stall forever). */
	if (avail < tableLen || avail < dataEnd) return 0;

	if (haveEncryption && (encryptionVal == 0x01 || encryptionVal == 0x03)) {
		/* ENCRYPT_ON / ENCRYPT_REQ: server requires TLS, which this
		 * library does not implement (see Common.h). */
		AltDB_DiagPushClient(slot, "08001", "server requires TLS encryption, not supported by this library");
		return -1;
	}

	c->TokPos += (tableLen > dataEnd) ? tableLen : dataEnd; /* consume exactly the parsed message */
	return 1;
}

/* ---------------- LOGIN7 ---------------- */

static UINT PutVarField(unsigned char *fixed, UINT pairOffset, unsigned char *var, UINT *varOff, UINT cap,
                         UINT encoding, const unsigned char *text, UDINT textLen)
{
	UINT chars;
	UDINT written;

	AltDB_WriteLE16(&fixed[pairOffset], (UINT)(94 + *varOff));
	written = AltDB_ConnToUtf16le(encoding, text, textLen, &var[*varOff], (cap > *varOff) ? (cap - *varOff) : 0);
	chars = (UINT)(written / 2);
	AltDB_WriteLE16(&fixed[pairOffset + 2], chars);
	*varOff += (UINT)written;
	return chars;
}

BOOL AltDB_BuildLogin7(UDINT slot, const char *user, const char *pass, const char *db, const char *server)
{
	ConnSlot *c = &gConn[slot];
	unsigned char *msg = c->SendBuf;
	unsigned char *fixed = &msg[8];
	unsigned char *var = &msg[8 + 94];
	UINT varCap = (UINT)(sizeof(c->SendBuf) - 8 - 94);
	UINT varOff = 0;
	UDINT total;
	UINT pwOff, pwChars, i;

	memset(msg, 0, sizeof(c->SendBuf));

	AltDB_WriteLE32(&fixed[4], 0x74000004UL);			/* TDSVersion 7.4 */
	AltDB_WriteLE32(&fixed[8], TDS_DEFAULT_PACKET_SIZE);	/* PacketSize */
	AltDB_WriteLE32(&fixed[12], 0x00010000UL);			/* ClientProgVer */
	AltDB_WriteLE32(&fixed[16], 0);						/* ClientPID */
	AltDB_WriteLE32(&fixed[20], 0);						/* ConnectionID */
	fixed[24] = 0xE0;										/* OptionFlags1 */
	fixed[25] = 0x03;										/* OptionFlags2 (fODBC=1) */
	fixed[26] = 0x00;										/* TypeFlags */
	fixed[27] = 0x00;										/* OptionFlags3 */
	AltDB_WriteLE32(&fixed[28], 0);						/* ClientTimeZone */
	AltDB_WriteLE32(&fixed[32], 0x00000409UL);			/* ClientLCID */

	PutVarField(fixed, 36, var, &varOff, varCap, c->Encoding, (const unsigned char *)"AltDB", 7); /* HostName */
	PutVarField(fixed, 40, var, &varOff, varCap, c->Encoding, (const unsigned char *)user, (UDINT)strlen(user)); /* UserName */

	pwOff = (UINT)(94 + varOff);
	pwChars = (UINT)(AltDB_ConnToUtf16le(c->Encoding, (const unsigned char *)pass, (UDINT)strlen(pass),
	                                        &var[varOff], varCap - varOff) / 2);
	for (i = 0; i < pwChars; i++) {
		unsigned char b0 = var[varOff + i * 2];
		unsigned char b1 = var[varOff + i * 2 + 1];
		b0 = (unsigned char)(((b0 << 4) | (b0 >> 4)) ^ 0xA5);
		b1 = (unsigned char)(((b1 << 4) | (b1 >> 4)) ^ 0xA5);
		var[varOff + i * 2] = b0;
		var[varOff + i * 2 + 1] = b1;
	}
	AltDB_WriteLE16(&fixed[44], pwOff);
	AltDB_WriteLE16(&fixed[46], pwChars);
	varOff += pwChars * 2;

	PutVarField(fixed, 48, var, &varOff, varCap, c->Encoding, (const unsigned char *)"AltDB", 7); /* AppName */
	PutVarField(fixed, 52, var, &varOff, varCap, c->Encoding, (const unsigned char *)server, (UDINT)strlen(server)); /* ServerName */
	AltDB_WriteLE16(&fixed[56], (UINT)(94 + varOff)); AltDB_WriteLE16(&fixed[58], 0); /* Extension: none */
	PutVarField(fixed, 60, var, &varOff, varCap, c->Encoding, (const unsigned char *)"AltDB", 7); /* CltIntName */
	AltDB_WriteLE16(&fixed[64], (UINT)(94 + varOff)); AltDB_WriteLE16(&fixed[66], 0); /* Language: none */
	PutVarField(fixed, 68, var, &varOff, varCap, c->Encoding, (const unsigned char *)db, (UDINT)strlen(db)); /* Database */

	memset(&fixed[72], 0, 6); /* ClientID */
	AltDB_WriteLE16(&fixed[78], (UINT)(94 + varOff)); AltDB_WriteLE16(&fixed[80], 0); /* SSPI: none */
	AltDB_WriteLE16(&fixed[82], (UINT)(94 + varOff)); AltDB_WriteLE16(&fixed[84], 0); /* AtchDBFile: none */
	AltDB_WriteLE16(&fixed[86], (UINT)(94 + varOff)); AltDB_WriteLE16(&fixed[88], 0); /* ChangePassword: none */
	AltDB_WriteLE32(&fixed[90], 0); /* cbSSPILong */

	total = 8 + 94 + varOff;
	AltDB_WriteLE32(&fixed[0], (UDINT)(94 + varOff));
	msg[0] = 0x10; msg[1] = 0x01; /* type LOGIN7, status EOM */
	AltDB_WriteBE16(&msg[2], (UINT)total);
	msg[4] = 0; msg[5] = 0; msg[6] = 1; msg[7] = 0;

	c->SendLen = total;
	c->SendPos = 0;
	return TRUE;
}

/* ---------------- SQL_BATCH (Section 10.6) ---------------- */

BOOL AltDB_BuildSqlBatch(UDINT slot, const char *sql, UDINT sqlLen)
{
	ConnSlot *c = &gConn[slot];
	unsigned char *msg = c->SendBuf;
	UDINT encCap = (UDINT)sizeof(c->SendBuf) - 8 - 22;
	UDINT encLen;
	UDINT total;

	encLen = AltDB_EncodeToWire(c->Encoding, sql, sqlLen, &msg[8 + 22], encCap);

	AltDB_WriteLE32(&msg[8 + 0], 22);		/* ALL_HEADERS TotalLength */
	AltDB_WriteLE32(&msg[8 + 4], 18);		/* HeaderLength */
	AltDB_WriteLE16(&msg[8 + 8], 2);			/* HeaderType: transaction descriptor */
	memcpy(&msg[8 + 10], c->TransactionDescr, 8);
	AltDB_WriteLE32(&msg[8 + 18], 1);		/* OutstandingRequestCount */

	total = 8 + 22 + encLen;
	msg[0] = 0x01; msg[1] = 0x01; /* type SQL_BATCH, status EOM */
	AltDB_WriteBE16(&msg[2], (UINT)total);
	msg[4] = 0; msg[5] = 0; msg[6] = 1; msg[7] = 0;

	c->SendLen = total;
	c->SendPos = 0;
	return TRUE;
}

/* ---------------- top level connect state machine ---------------- */

INT AltDB_NetConnectStep(UDINT slot)
{
	ConnSlot *c = &gConn[slot];
	INT r;

	switch (c->State) {

	case CONNSTATE_OPENING:
		r = PumpTcpOpen(slot);
		if (r == NET_IN_PROGRESS) return NET_IN_PROGRESS;
		if (r == NET_ERROR) { c->State = CONNSTATE_FAILED; return NET_ERROR; }
		c->State = CONNSTATE_CONNECTING;
		return NET_IN_PROGRESS;

	case CONNSTATE_CONNECTING:
		r = PumpTcpClient(slot);
		if (r == NET_IN_PROGRESS) return NET_IN_PROGRESS;
		if (r == NET_ERROR) { c->State = CONNSTATE_FAILED; return NET_ERROR; }
		c->State = CONNSTATE_PRELOGIN;
		c->NetStep = NETSTEP_SEND;
		AltDB_BuildPrelogin(slot);
		return NET_IN_PROGRESS;

	case CONNSTATE_PRELOGIN:
		if (c->NetStep == NETSTEP_SEND) {
			r = AltDB_NetSendStep(slot);
			if (r == NET_ERROR) { c->State = CONNSTATE_FAILED; return NET_ERROR; }
			if (r == NET_DONE) c->NetStep = NETSTEP_RECV;
			return NET_IN_PROGRESS;
		} else {
			r = AltDB_NetRecvPump(slot);
			if (r < 0) { c->State = CONNSTATE_FAILED; return NET_ERROR; }
			r = ParsePreloginResponse(slot);
			if (r < 0) { c->State = CONNSTATE_FAILED; return NET_ERROR; }
			if (r == 0) return NET_IN_PROGRESS;
			/* ParsePreloginResponse already advanced TokPos past exactly
			 * the bytes it consumed; nothing is discarded here. */
			c->State = CONNSTATE_LOGIN;
			c->NetStep = NETSTEP_SEND;
			AltDB_BuildLogin7(slot, (const char *)c->LoginUser, (const char *)c->LoginPass,
			                    (const char *)c->LoginDb, (const char *)c->HostBuf);
			return NET_IN_PROGRESS;
		}

	case CONNSTATE_LOGIN:
		if (c->NetStep == NETSTEP_SEND) {
			r = AltDB_NetSendStep(slot);
			if (r == NET_ERROR) { c->State = CONNSTATE_FAILED; return NET_ERROR; }
			if (r == NET_DONE) c->NetStep = NETSTEP_RECV;
			return NET_IN_PROGRESS;
		} else {
			INT tok;
			r = AltDB_NetRecvPump(slot);
			if (r < 0) { c->State = CONNSTATE_FAILED; return NET_ERROR; }
			tok = AltDB_TokenStep(slot, TOKMODE_LOGIN);
			if (tok == TOK_NEED_MORE) return NET_IN_PROGRESS;
			if (tok == TOK_ERROR) { c->State = CONNSTATE_FAILED; return NET_ERROR; }
			/* TOK_GOT_DONE_FINAL: login succeeded */
			c->State = CONNSTATE_IDLE;
			return NET_DONE;
		}

	default:
		return NET_ERROR;
	}
}
```

#### Token.c - TDS response token stream parser
```c
/********************************************************************
 * Library: AltDB
 * File: Token.c
 ********************************************************************
 * Incremental TDS response token stream parser (Section 10.7). Reads
 * from gConn[slot].TokBuf[TokPos..TokLen) which already has the
 * 8-byte TDS packet headers stripped (Net.c). Never blocks: if a
 * token is not yet fully buffered, parsing stops without consuming
 * it and is resumed transparently on the next call once more bytes
 * have arrived - the parser carries no state beyond (TokBuf, TokPos).
 ********************************************************************/
#include <bur/plctypes.h>
#include <runtime.h>
#include <AsTCP.h>
#include <AltDB.h>
#include "Common.h"
#include <string.h>

/* TDS type ids (Section 10.9 / Table 21) */
#define TY_NULL        0x1F
#define TY_INT1        0x30
#define TY_BIT         0x32
#define TY_INT2        0x34
#define TY_INT4        0x38
#define TY_DATETIM4    0x3A
#define TY_FLT4        0x3B
#define TY_MONEY       0x3C
#define TY_DATETIME    0x3D
#define TY_FLT8        0x3E
#define TY_MONEY4      0x7A
#define TY_INT8        0x7F
#define TY_INTN        0x26
#define TY_BITN        0x68
#define TY_FLTN        0x6D
#define TY_MONEYN      0x6E
#define TY_DATETIMN    0x6F
#define TY_GUID        0x24
#define TY_DECIMALN    0x6A
#define TY_NUMERICN    0x6C
#define TY_DATEN       0x28
#define TY_TIMEN       0x29
#define TY_DATETIME2N  0x2A
#define TY_DATETIMEOFFSETN 0x2B
#define TY_BIGVARCHR   0xA7
#define TY_BIGCHAR     0xAF
#define TY_NVARCHAR    0xE7
#define TY_NCHAR       0xEF
#define TY_BIGVARBIN   0xA5
#define TY_BIGBINARY   0xAD
#define TY_CHAR_LEGACY     0x2F
#define TY_VARCHAR_LEGACY  0x27
#define TY_BINARY_LEGACY   0x2D
#define TY_VARBINARY_LEGACY 0x25
#define TY_TEXT        0x23
#define TY_NTEXT       0x63
#define TY_IMAGE       0x22
#define TY_VARIANT     0x62
#define TY_XML         0xF1
#define TY_UDT         0xF0

/* ---------------- TYPE_INFO parsing (COLMETADATA) ---------------- */

/* Returns bytes of TYPE_INFO consumed (>=1), 0 if more bytes are
 * needed, -1 if the type byte is not a recognised TDS data type
 * (unrecoverable: we cannot safely determine its size). */
static INT ParseTypeInfo(const unsigned char *b, UDINT avail, ColumnInfo *col)
{
	UDINT pos = 1;
	unsigned char t;

	if (avail < 1) return 0;
	t = b[0];
	col->DataType = t;
	col->IsUnicode = FALSE;
	col->IsPlp = FALSE;
	col->IsLongLen = FALSE;
	col->Supported = TRUE;
	col->Precision = 0;
	col->Scale = 0;
	col->MaxLength = 0;

	switch (t) {
	case TY_NULL:
		col->MaxLength = 0;
		break;
	case TY_INT1: case TY_BIT:
		col->MaxLength = 1;
		break;
	case TY_INT2:
		col->MaxLength = 2;
		break;
	case TY_INT4: case TY_DATETIM4: case TY_FLT4: case TY_MONEY4:
		col->MaxLength = 4;
		break;
	case TY_MONEY: case TY_DATETIME: case TY_FLT8: case TY_INT8:
		col->MaxLength = 8;
		break;

	case TY_INTN: case TY_BITN: case TY_FLTN: case TY_MONEYN: case TY_DATETIMN: case TY_GUID:
		if (avail < pos + 1) return 0;
		col->MaxLength = b[pos]; pos += 1;
		break;

	case TY_DECIMALN: case TY_NUMERICN:
		if (avail < pos + 3) return 0;
		col->MaxLength = b[pos]; col->Precision = b[pos + 1]; col->Scale = b[pos + 2];
		pos += 3;
		break;

	case TY_DATEN:
		break; /* no extra TYPE_INFO byte */
	case TY_TIMEN: case TY_DATETIME2N: case TY_DATETIMEOFFSETN:
		if (avail < pos + 1) return 0;
		col->Scale = b[pos]; pos += 1;
		break;

	case TY_BIGVARCHR: case TY_BIGCHAR: case TY_NVARCHAR: case TY_NCHAR:
	case TY_BIGVARBIN: case TY_BIGBINARY: {
		UINT maxLen;
		if (avail < pos + 2) return 0;
		maxLen = (UINT)AltDB_ReadLE16(&b[pos]); pos += 2;
		col->MaxLength = maxLen;
		col->IsPlp = (maxLen == 0xFFFF);
		col->IsUnicode = (t == TY_NVARCHAR || t == TY_NCHAR);
		if (t == TY_BIGVARCHR || t == TY_BIGCHAR || t == TY_NVARCHAR || t == TY_NCHAR) {
			if (avail < pos + 5) return 0;
			pos += 5; /* collation, not required for the supported conversions */
		}
		break;
	}

	case TY_CHAR_LEGACY: case TY_VARCHAR_LEGACY: case TY_BINARY_LEGACY: case TY_VARBINARY_LEGACY:
		if (avail < pos + 1) return 0;
		col->MaxLength = b[pos]; pos += 1;
		break;

	case TY_TEXT: case TY_NTEXT: case TY_IMAGE: {
		UDINT i;
		unsigned char numParts;
		if (avail < pos + 4) return 0;
		col->MaxLength = AltDB_ReadLE32(&b[pos]); pos += 4;
		col->IsLongLen = TRUE;
		col->IsUnicode = (t == TY_NTEXT);
		if (t != TY_IMAGE) {
			if (avail < pos + 5) return 0;
			pos += 5; /* collation */
		}
		if (avail < pos + 1) return 0;
		numParts = b[pos]; pos += 1;
		for (i = 0; i < numParts; i++) {
			UINT n;
			if (avail < pos + 2) return 0;
			n = (UINT)AltDB_ReadLE16(&b[pos]);
			if (avail < pos + 2 + (UDINT)n * 2) return 0;
			pos += 2 + (UDINT)n * 2;
		}
		break;
	}

	case TY_VARIANT:
		if (avail < pos + 4) return 0;
		col->MaxLength = AltDB_ReadLE32(&b[pos]); pos += 4;
		col->Supported = FALSE;
		break;

	case TY_XML: {
		unsigned char schemaPresent;
		if (avail < pos + 1) return 0;
		schemaPresent = b[pos]; pos += 1;
		col->IsPlp = TRUE;
		col->IsUnicode = TRUE;
		col->Supported = FALSE;
		if (schemaPresent) {
			UDINT i;
			for (i = 0; i < 3; i++) {
				UDINT n;
				if (i < 2) {
					if (avail < pos + 1) return 0;
					n = b[pos]; pos += 1;
				} else {
					if (avail < pos + 2) return 0;
					n = AltDB_ReadLE16(&b[pos]); pos += 2;
				}
				if (avail < pos + n * 2) return 0;
				pos += n * 2;
			}
		}
		break;
	}

	case TY_UDT: {
		UDINT i;
		if (avail < pos + 2) return 0;
		pos += 2; /* MAX_BYTE_SIZE */
		col->IsPlp = TRUE;
		col->Supported = FALSE;
		for (i = 0; i < 4; i++) {
			UDINT n;
			if (i < 3) { /* DB_NAME, SCHEMA_NAME, TYPE_NAME: B_VARCHAR */
				if (avail < pos + 1) return 0;
				n = b[pos]; pos += 1;
			} else { /* ASSEMBLY_QUALIFIED_NAME: US_VARCHAR */
				if (avail < pos + 2) return 0;
				n = AltDB_ReadLE16(&b[pos]); pos += 2;
			}
			if (avail < pos + n * 2) return 0;
			pos += n * 2;
		}
		break;
	}

	default:
		return -1;
	}

	return (INT)pos;
}

/* TRUE for byte-length-class types whose value carries a 1-byte
 * length prefix with 0 meaning NULL (as opposed to legal zero-length
 * non-NULL content). */
static BOOL IsByteLenNullable(unsigned char t)
{
	switch (t) {
	case TY_INTN: case TY_BITN: case TY_FLTN: case TY_MONEYN: case TY_DATETIMN: case TY_GUID:
	case TY_DECIMALN: case TY_NUMERICN:
	case TY_DATEN: case TY_TIMEN: case TY_DATETIME2N: case TY_DATETIMEOFFSETN:
		return TRUE;
	default:
		return FALSE;
	}
}

/* Parses one column value from the ROW/NBCROW wire format into dst
 * (clamped to dstCap; *outValLen reports the true, unclamped length
 * so overflow can be detected by the caller). Returns bytes consumed
 * from the wire (>0), 0 if more bytes are needed, -1 on a malformed
 * value that cannot be safely skipped. */
static INT ParseColumnValue(const unsigned char *b, UDINT avail, const ColumnInfo *col,
                             unsigned char *dst, UDINT dstCap, UDINT *outValLen, BOOL *outIsNull)
{
	unsigned char t = col->DataType;
	UDINT fixedLen = 0;

	*outValLen = 0;
	*outIsNull = FALSE;

	switch (t) {
	case TY_NULL: *outIsNull = TRUE; return 0;
	case TY_INT1: case TY_BIT: fixedLen = 1; break;
	case TY_INT2: fixedLen = 2; break;
	case TY_INT4: case TY_DATETIM4: case TY_FLT4: case TY_MONEY4: fixedLen = 4; break;
	case TY_MONEY: case TY_DATETIME: case TY_FLT8: case TY_INT8: fixedLen = 8; break;
	default: fixedLen = 0; break;
	}

	if (fixedLen > 0) {
		if (avail < fixedLen) return 0;
		*outValLen = fixedLen;
		memcpy(dst, b, (fixedLen < dstCap) ? fixedLen : dstCap);
		return (INT)fixedLen;
	}

	if (col->IsPlp) {
		/* PLP (Section 10.9): 8-byte total length, then chunks of
		 * (4-byte length, data), terminated by a 4-byte zero length.
		 * 0xFFFFFFFFFFFFFFFF total length = NULL. */
		unsigned long long total;
		UDINT pos = 8;
		UDINT copied = 0;

		if (avail < 8) return 0;
		total = AltDB_ReadLE64(b);
		if (total == 0xFFFFFFFFFFFFFFFFULL) { *outIsNull = TRUE; return 8; }

		for (;;) {
			UDINT chunkLen;
			if (avail < pos + 4) return 0;
			chunkLen = AltDB_ReadLE32(&b[pos]); pos += 4;
			if (chunkLen == 0) break;
			if (avail < pos + chunkLen) return 0;
			if (copied < dstCap) {
				UDINT n = chunkLen;
				if (copied + n > dstCap) n = dstCap - copied;
				memcpy(&dst[copied], &b[pos], n);
			}
			copied += chunkLen;
			pos += chunkLen;
		}
		*outValLen = copied;
		return (INT)pos;
	}

	if (col->IsLongLen) {
		/* Legacy TEXT/NTEXT/IMAGE: 1-byte TEXTPTR length (0 = NULL),
		 * TEXTPTR bytes, 8-byte timestamp, 4-byte data length, data. */
		UDINT pos = 0;
		unsigned char ptrLen;

		if (avail < 1) return 0;
		ptrLen = b[0]; pos = 1;
		if (ptrLen == 0) { *outIsNull = TRUE; return (INT)pos; }
		if (avail < pos + ptrLen + 8 + 4) return 0;
		pos += ptrLen + 8;
		{
			UDINT dataLen = AltDB_ReadLE32(&b[pos]); pos += 4;
			if (avail < pos + dataLen) return 0;
			*outValLen = dataLen;
			memcpy(dst, &b[pos], (dataLen < dstCap) ? dataLen : dstCap);
			pos += dataLen;
			return (INT)pos;
		}
	}

	if (t == TY_VARIANT) {
		UDINT total;
		if (avail < 4) return 0;
		total = AltDB_ReadLE32(b);
		if (total == 0) { *outIsNull = TRUE; return 4; }
		if (avail < 4 + total) return 0;
		/* BaseType + PropBytes + Value; copy raw for completeness, not
		 * decoded further (col->Supported is FALSE for SQL_VARIANT). */
		*outValLen = total;
		memcpy(dst, &b[4], (total < dstCap) ? total : dstCap);
		return (INT)(4 + total);
	}

	if (IsByteLenNullable(t)) {
		UDINT len;
		if (avail < 1) return 0;
		len = b[0];
		if (len == 0) { *outIsNull = TRUE; return 1; }
		if (avail < 1 + len) return 0;
		*outValLen = len;
		memcpy(dst, &b[1], (len < dstCap) ? len : dstCap);
		return (INT)(1 + len);
	}

	switch (t) {
	case TY_BIGVARCHR: case TY_BIGCHAR: case TY_NVARCHAR: case TY_NCHAR:
	case TY_BIGVARBIN: case TY_BIGBINARY: {
		UDINT len;
		if (avail < 2) return 0;
		len = AltDB_ReadLE16(b);
		if (len == 0xFFFF) { *outIsNull = TRUE; return 2; }
		if (avail < 2 + len) return 0;
		*outValLen = len;
		memcpy(dst, &b[2], (len < dstCap) ? len : dstCap);
		return (INT)(2 + len);
	}
	case TY_CHAR_LEGACY: case TY_VARCHAR_LEGACY: case TY_BINARY_LEGACY: case TY_VARBINARY_LEGACY: {
		UDINT len;
		if (avail < 1) return 0;
		len = b[0];
		if (avail < 1 + len) return 0;
		*outValLen = len; /* legacy types have no dedicated NULL sentinel here */
		memcpy(dst, &b[1], (len < dstCap) ? len : dstCap);
		return (INT)(1 + len);
	}
	default:
		return -1;
	}
}

/* ---------------- COLMETADATA (0x81) ---------------- */

static INT ParseColMetadata(UDINT slot)
{
	ConnSlot *c = &gConn[slot];
	const unsigned char *b = &c->TokBuf[c->TokPos];
	UDINT avail = c->TokLen - c->TokPos;
	UDINT pos = 1;
	UINT count;
	UINT colIdx;
	ColumnInfo overflowCol;

	if (avail < 3) return 0;
	count = (UINT)AltDB_ReadLE16(&b[1]);
	pos = 3;
	if (count == 0xFFFF) count = 0;

	for (colIdx = 0; colIdx < count; colIdx++) {
		ColumnInfo *dst = (colIdx < ND_MAX_COLUMNS) ? &c->Columns[colIdx] : &overflowCol;
		INT tiLen;
		UINT nameLen;

		if (avail < pos + 6) return 0; /* UserType(4) + Flags(2) */
		pos += 6;

		tiLen = ParseTypeInfo(&b[pos], avail - pos, dst);
		if (tiLen == 0) return 0;
		if (tiLen < 0) { AltDB_DiagPushClient(slot, "HY000", "unrecognised TDS column type"); return -1; }
		pos += (UDINT)tiLen;

		if (avail < pos + 1) return 0;
		nameLen = b[pos];
		if (avail < pos + 1 + (UDINT)nameLen * 2) return 0;
		pos += 1 + (UDINT)nameLen * 2;
	}

	c->ColumnCount = (count > 0x7FFF) ? 0x7FFF : (INT)count;
	memset(c->ColAlreadyRead, 0, sizeof(c->ColAlreadyRead));
	memset(c->ColIsNull, 0, sizeof(c->ColIsNull));
	c->RowReady = FALSE;
	c->RowOverflow = FALSE;
	c->HasResultSet = TRUE;
	c->ResultSetOpen = TRUE;
	c->TokPos += pos;
	return 1;
}

/* ---------------- ROW (0xD1) / NBCROW (0xD2) ---------------- */

static INT ParseRow(UDINT slot, BOOL isNbc)
{
	ConnSlot *c = &gConn[slot];
	const unsigned char *b = &c->TokBuf[c->TokPos];
	UDINT avail = c->TokLen - c->TokPos;
	UDINT pos = 1;
	INT colCount = (c->ColumnCount > 0) ? c->ColumnCount : 0;
	UDINT nullBitmapBytes = 0;
	const unsigned char *nullBitmap = NULL;
	INT i;
	BOOL overflow = FALSE;

	if (isNbc) {
		nullBitmapBytes = ((UDINT)colCount + 7) / 8;
		if (avail < pos + nullBitmapBytes) return 0;
		nullBitmap = &b[pos];
		pos += nullBitmapBytes;
	}

	for (i = 0; i < colCount; i++) {
		BOOL bitmapNull = FALSE;
		BOOL isNull = FALSE;
		UDINT valLen = 0;
		INT consumed;
		ColumnInfo dummyCol;
		ColumnInfo *col;
		unsigned char dummyDst[1];
		unsigned char *dst;
		UDINT dstCap;

		if (isNbc && (nullBitmap[i / 8] & (1 << (i % 8))) != 0) {
			bitmapNull = TRUE;
		}

		if (i < ND_MAX_COLUMNS) {
			col = &c->Columns[i];
			dst = c->ColValue[i];
			dstCap = ND_MAX_COL_VALUE_LEN;
		} else {
			/* Columns beyond ND_MAX_COLUMNS: metadata was not retained
			 * (ParseColMetadata), so the value cannot be decoded. This
			 * is only reachable for results with more columns than
			 * this library supports and is reported as dbERR_MEMORY
			 * by the caller via RowOverflow. */
			memset(&dummyCol, 0, sizeof(dummyCol));
			dummyCol.DataType = TY_NULL;
			col = &dummyCol;
			dst = dummyDst;
			dstCap = 0;
			overflow = TRUE;
		}

		if (bitmapNull) {
			isNull = TRUE;
			consumed = 0;
		} else {
			consumed = ParseColumnValue(&b[pos], avail - pos, col, dst, dstCap, &valLen, &isNull);
			if (consumed == 0) return 0;
			if (consumed < 0) { AltDB_DiagPushClient(slot, "HY000", "malformed row value"); return -1; }
		}
		pos += (UDINT)consumed;

		if (i < ND_MAX_COLUMNS) {
			c->ColIsNull[i] = isNull;
			c->ColAlreadyRead[i] = FALSE;
			if (!isNull) {
				c->ColValueLen[i] = valLen;
				if (valLen > ND_MAX_COL_VALUE_LEN) overflow = TRUE;
			} else {
				c->ColValueLen[i] = 0;
			}
		}
	}

	c->TokPos += pos;
	c->RowReady = TRUE;
	c->RowOverflow = overflow;
	return 1;
}

/* ---------------- ERROR (0xAA) / INFO (0xAB) ---------------- */

static void MapSqlState(DINT nativeError, unsigned char class_, BOOL isError, char out[6])
{
	const char *s;

	if (!isError) { s = "01000"; }
	else switch (nativeError) {
		case 18456: s = "28000"; break;
		case 4060:  s = "42000"; break;
		case 102: case 156: s = "42000"; break;
		case 208: s = "42S02"; break;
		case 207: s = "42S22"; break;
		case 2627: case 2601: case 547: case 515: s = "23000"; break;
		case 8152: case 2628: s = "22001"; break;
		case 245: case 8114: s = "22018"; break;
		case 8115: s = "22003"; break;
		case 1205: s = "40001"; break;
		default: s = (class_ >= 17) ? "HY000" : "42000"; break;
	}
	memcpy(out, s, 5);
	out[5] = 0;
}

static INT ParseErrorOrInfo(UDINT slot, BOOL isError)
{
	ConnSlot *c = &gConn[slot];
	const unsigned char *b = &c->TokBuf[c->TokPos];
	UDINT avail = c->TokLen - c->TokPos;
	UINT length;
	UDINT total;
	DINT number;
	unsigned char class_;
	UINT msgChars;
	UDINT msgBytes;
	char sqlState[6];
	unsigned char connMsg[256];
	UDINT connMsgLen;

	if (avail < 3) return 0;
	length = (UINT)AltDB_ReadLE16(&b[1]);
	total = 3 + length;
	if (avail < total) return 0;

	number = (DINT)AltDB_ReadLE32(&b[3]);
	/* b[7] = State (1 byte), b[8] = Class (1 byte) */
	class_ = b[8];
	msgChars = (UINT)AltDB_ReadLE16(&b[9]);
	msgBytes = (UDINT)msgChars * 2;

	MapSqlState(number, class_, isError && class_ >= 11, sqlState);
	connMsgLen = AltDB_WireToConn(c->Encoding, &b[11], msgBytes, connMsg, sizeof(connMsg));
	AltDB_DiagPushServer(slot, isError && class_ >= 11, number, sqlState, connMsg, connMsgLen);

	c->TokPos += total;
	return 1;
}

/* ---------------- LOGINACK (0xAD) ---------------- */

static INT ParseLoginAck(UDINT slot)
{
	ConnSlot *c = &gConn[slot];
	const unsigned char *b = &c->TokBuf[c->TokPos];
	UDINT avail = c->TokLen - c->TokPos;
	UINT length;
	UDINT total;

	if (avail < 3) return 0;
	length = (UINT)AltDB_ReadLE16(&b[1]);
	total = 3 + length;
	if (avail < total) return 0;

	if (length >= 10) {
		/* payload (offset 3 = start of token data): Interface(1) at 3,
		 * TDSVersion(4) at 4..7, ProgName B_VARCHAR length byte at 8,
		 * ProgName chars at 9.., ProgVersion(4) right after. */
		UDINT progNameLenPos = 8;
		UINT progNameChars = b[progNameLenPos];
		UDINT progVerPos = progNameLenPos + 1 + (UDINT)progNameChars * 2;

		if (avail >= progVerPos + 4) {
			unsigned char major = b[progVerPos];
			unsigned char minor = b[progVerPos + 1];
			UINT build = (UINT)((b[progVerPos + 2] << 8) | b[progVerPos + 3]);
			char tmp[32];
			UDINT n = 0;

			n += AltDB_FormatI64(major, &tmp[n], sizeof(tmp) - n);
			tmp[n++] = '.';
			n += AltDB_FormatI64(minor, &tmp[n], sizeof(tmp) - n);
			tmp[n++] = '.';
			n += AltDB_FormatI64(build, &tmp[n], sizeof(tmp) - n);
			if (n >= sizeof(c->ServerVersion)) n = sizeof(c->ServerVersion) - 1;
			memcpy(c->ServerVersion, tmp, n);
			c->ServerVersion[n] = 0;
		}
	}

	c->TokPos += total;
	return 1;
}

/* ---------------- ENVCHANGE (0xE3) ---------------- */

static INT ParseEnvChange(UDINT slot)
{
	ConnSlot *c = &gConn[slot];
	const unsigned char *b = &c->TokBuf[c->TokPos];
	UDINT avail = c->TokLen - c->TokPos;
	UINT length;
	UDINT total;
	unsigned char envType;

	if (avail < 3) return 0;
	length = (UINT)AltDB_ReadLE16(&b[1]);
	total = 3 + length;
	if (avail < total) return 0;

	envType = (length >= 1) ? b[3] : 0;

	if (envType == 4 && length >= 2) {
		/* packet size: NewValue is a B_VARCHAR of decimal digit characters */
		UINT nChars = b[4];
		UDINT i;
		UDINT v = 0;
		for (i = 0; i < nChars && (5 + i * 2 + 1) < total; i++) {
			unsigned char ch = b[5 + i * 2];
			if (ch >= '0' && ch <= '9') v = v * 10 + (UDINT)(ch - '0');
		}
		if (v > 0 && v <= 32768) c->PacketSize = (UINT)v;
	} else if ((envType == 8 || envType == 9 || envType == 10 || envType == 17) && length >= 2) {
		unsigned char n = b[4];
		if (n == 8 && total >= 5 + 8) {
			memcpy(c->TransactionDescr, &b[5], 8);
		}
	}

	c->TokPos += total;
	return 1;
}

/* ---------------- generic Length-prefixed skip ---------------- */

static INT SkipLengthPrefixed16(UDINT slot)
{
	ConnSlot *c = &gConn[slot];
	const unsigned char *b = &c->TokBuf[c->TokPos];
	UDINT avail = c->TokLen - c->TokPos;
	UINT length;

	if (avail < 3) return 0;
	length = (UINT)AltDB_ReadLE16(&b[1]);
	if (avail < (UDINT)(3 + length)) return 0;
	c->TokPos += 3 + length;
	return 1;
}

static INT SkipSessionState(UDINT slot)
{
	ConnSlot *c = &gConn[slot];
	const unsigned char *b = &c->TokBuf[c->TokPos];
	UDINT avail = c->TokLen - c->TokPos;
	UDINT length;

	if (avail < 5) return 0;
	length = AltDB_ReadLE32(&b[1]);
	if (avail < 5 + length) return 0;
	c->TokPos += 5 + length;
	return 1;
}

/* ---------------- DONE / DONEPROC / DONEINPROC (0xFD/0xFE/0xFF) ---------------- */

#define DONE_MORE     0x0001
#define DONE_ERROR    0x0002
#define DONE_COUNT    0x0010
#define DONE_SRVERROR 0x0100

static INT ParseDone(UDINT slot, BOOL *outMore, BOOL *outError)
{
	ConnSlot *c = &gConn[slot];
	const unsigned char *b = &c->TokBuf[c->TokPos];
	UDINT avail = c->TokLen - c->TokPos;
	UINT status;
	unsigned long long rowCount;

	if (avail < 13) return 0;
	status = (UINT)AltDB_ReadLE16(&b[1]);
	rowCount = AltDB_ReadLE64(&b[5]);

	*outMore = (status & DONE_MORE) != 0;
	*outError = (status & (DONE_ERROR | DONE_SRVERROR)) != 0;

	if ((status & DONE_COUNT) != 0 && !c->AffectedRowsKnown) {
		c->AffectedRows = (rowCount > 0xFFFFFFFFULL) ? 0xFFFFFFFFUL : (UDINT)rowCount;
		c->AffectedRowsKnown = TRUE;
	}

	c->TokPos += 13;
	return 1;
}

/* ---------------- top level dispatcher ---------------- */

INT AltDB_TokenStep(UDINT slot, UINT mode)
{
	ConnSlot *c = &gConn[slot];
	BOOL sawError = FALSE;

	for (;;) {
		unsigned char tokType;
		INT r;

		if (c->TokPos >= c->TokLen) return TOK_NEED_MORE;
		tokType = c->TokBuf[c->TokPos];

		switch (tokType) {
		case 0x81: /* COLMETADATA */
			r = ParseColMetadata(slot);
			if (r == 0) return TOK_NEED_MORE;
			if (r < 0) return TOK_ERROR;
			if (mode == TOKMODE_EXEC) return TOK_GOT_COLMETADATA;
			/* FETCH/DRAIN: a later statement's columns; keep consuming */
			break;

		case 0xD1: /* ROW */
		case 0xD2: /* NBCROW */
			r = ParseRow(slot, (tokType == 0xD2));
			if (r == 0) return TOK_NEED_MORE;
			if (r < 0) return TOK_ERROR;
			if (c->RowOverflow) return TOK_ERROR_MEMORY;
			if (mode == TOKMODE_FETCH) return TOK_GOT_ROW;
			/* EXEC should not normally see rows before COLMETADATA is
			 * returned to the caller; DRAIN discards them. */
			break;

		case 0xFD: case 0xFE: case 0xFF: { /* DONE / DONEPROC / DONEINPROC */
			BOOL more, errFlag;
			r = ParseDone(slot, &more, &errFlag);
			if (r == 0) return TOK_NEED_MORE;

			if (mode == TOKMODE_FETCH) {
				c->ResultSetOpen = FALSE;
				c->NoMoreRows = TRUE;
				return (errFlag || sawError) ? TOK_ERROR : TOK_GOT_EOF;
			}
			if (errFlag || sawError) return TOK_ERROR;
			if (more) break; /* more statements follow in this batch */
			if (mode == TOKMODE_DRAIN) return TOK_GOT_DONE_FINAL;
			if (mode == TOKMODE_LOGIN) return TOK_GOT_DONE_FINAL;
			/* TOKMODE_EXEC: batch ended without ever producing a result set */
			c->HasResultSet = FALSE;
			c->ResultSetOpen = FALSE;
			return TOK_GOT_DONE_FINAL;
		}

		case 0xAA: /* ERROR */
			r = ParseErrorOrInfo(slot, TRUE);
			if (r == 0) return TOK_NEED_MORE;
			sawError = TRUE;
			break;

		case 0xAB: /* INFO */
			r = ParseErrorOrInfo(slot, FALSE);
			if (r == 0) return TOK_NEED_MORE;
			break;

		case 0xAD: /* LOGINACK */
			r = ParseLoginAck(slot);
			if (r == 0) return TOK_NEED_MORE;
			break;

		case 0xE3: /* ENVCHANGE */
			r = ParseEnvChange(slot);
			if (r == 0) return TOK_NEED_MORE;
			break;

		case 0x79: /* RETURNSTATUS: fixed 4-byte value, ignored */
			if (c->TokLen - c->TokPos < 5) return TOK_NEED_MORE;
			c->TokPos += 5;
			break;

		case 0xA9: /* ORDER */
		case 0xA4: /* TABNAME */
		case 0xA5: /* COLINFO */
			r = SkipLengthPrefixed16(slot);
			if (r == 0) return TOK_NEED_MORE;
			break;

		case 0xE4: /* SESSIONSTATE */
			r = SkipSessionState(slot);
			if (r == 0) return TOK_NEED_MORE;
			break;

		default:
			AltDB_DiagPushClient(slot, "08S01", "unexpected/unsupported TDS token, protocol out of sync");
			return TOK_ERROR;
		}
	}
}
```
